  MoveL 2827 to (-200, -40.67, 52.07) mm, rotated rx 123.54 ry 0 rz 180 deg; joints [-9.323, -80.006, 124.061, 166.716, 44.832, -136.951]
  MoveL 2828 to (0, -40.67, 52.07) mm, rotated rx 123.54 ry 0 rz 180 deg; joints [-7.983, -68.226, 108.402, 167.736, 40.83, -137.116]
  MoveL 2829 to (0, -40.33, 52.56) mm, rotated rx 126.23 ry 0 rz 180 deg; joints [-8.518, -67.714, 108.589, 167.109, 41.6, -134.058]
  MoveL 2830 to (-200, -40.33, 52.56) mm, rotated rx 126.23 ry 0 rz 180 deg; joints [-9.945, -79.388, 124.274, 166.047, 45.743, -133.933]
  MoveL 2831 to (-200, -39.96, 53.04) mm, rotated rx 128.92 ry 0 rz 180 deg; joints [-10.538, -78.733, 124.49, 165.444, 46.691, -130.985]
  MoveL 2832 to (0, -39.96, 53.04) mm, rotated rx 128.92 ry 0 rz 180 deg; joints [-9.029, -67.172, 108.78, 166.542, 42.401, -131.062]
  MoveL 2833 to (0, -39.57, 53.5) mm, rotated rx 131.6 ry 0 rz 180 deg; joints [-9.515, -66.6, 108.972, 166.034, 43.23, -128.128]
  MoveL 2834 to (-200, -39.57, 53.5) mm, rotated rx 131.6 ry 0 rz 180 deg; joints [-11.101, -78.04, 124.71, 164.904, 47.673, -128.104]
  MoveL 2835 to (-200, -39.16, 53.94) mm, rotated rx 134.29 ry 0 rz 180 deg; joints [-11.634, -77.311, 124.93, 164.426, 48.684, -125.287]
  MoveL 2836 to (0, -39.16, 53.94) mm, rotated rx 134.29 ry 0 rz 180 deg; joints [-9.975, -65.998, 109.167, 165.583, 44.084, -125.251]
  MoveL 2837 to (0, -38.73, 54.36) mm, rotated rx 136.97 ry 0 rz 180 deg; joints [-10.407, -65.369, 109.361, 165.188, 44.96, -122.429]
  MoveL 2838 to (-200, -38.73, 54.36) mm, rotated rx 136.97 ry 0 rz 180 deg; joints [-12.134, -76.548, 125.152, 164.007, 49.723, -122.53]
  MoveL 2839 to (-200, -38.29, 54.76) mm, rotated rx 139.66 ry 0 rz 180 deg; joints [-12.602, -75.751, 125.373, 163.644, 50.786, -119.831]
  MoveL 2840 to (0, -38.29, 54.76) mm, rotated rx 139.66 ry 0 rz 180 deg; joints [-10.812, -64.712, 109.555, 164.846, 45.857, -119.661]
  MoveL 2841 to (0, -37.82, 55.13) mm, rotated rx 142.34 ry 0 rz 180 deg; joints [-11.188, -64.03, 109.748, 164.556, 46.771, -116.941]
  MoveL 2842 to (-200, -37.82, 55.13) mm, rotated rx 142.34 ry 0 rz 180 deg; joints [-13.037, -74.922, 125.593, 163.335, 51.871, -117.184]
  MoveL 2843 to (-200, -37.34, 55.49) mm, rotated rx 145.03 ry 0 rz 180 deg; joints [-13.438, -74.063, 125.81, 163.077, 52.974, -114.588]
  MoveL 2844 to (0, -37.34, 55.49) mm, rotated rx 145.03 ry 0 rz 180 deg; joints [-11.536, -63.323, 109.939, 164.314, 47.701, -114.267]
  MoveL 2845 to (0, -36.84, 55.82) mm, rotated rx 147.72 ry 0 rz 180 deg; joints [-11.853, -62.592, 110.127, 164.118, 48.643, -111.637]
  MoveL 2846 to (-200, -36.84, 55.82) mm, rotated rx 147.72 ry 0 rz 180 deg; joints [-13.804, -73.174, 126.025, 162.868, 54.095, -112.037]
  MoveL 2847 to (-200, -36.32, 56.13) mm, rotated rx 150.4 ry 0 rz 180 deg; joints [-14.135, -72.258, 126.235, 162.705, 55.228, -109.53]
  MoveL 2848 to (0, -36.32, 56.13) mm, rotated rx 150.4 ry 0 rz 180 deg; joints [-12.14, -61.84, 110.312, 163.968, 49.597, -109.048]
  MoveL 2849 to (0, -35.79, 56.41) mm, rotated rx 153.09 ry 0 rz 180 deg; joints [-12.397, -61.067, 110.492, 163.86, 50.559, -106.496]
  MoveL 2850 to (-200, -35.79, 56.41) mm, rotated rx 153.09 ry 0 rz 180 deg; joints [-14.43, -71.315, 126.439, 162.585, 56.374, -107.059]
  MoveL 2851 to (-200, -35.25, 56.67) mm, rotated rx 155.77 ry 0 rz 180 deg; joints [-14.69, -70.349, 126.638, 162.508, 57.53, -104.624]
  MoveL 2852 to (0, -35.25, 56.67) mm, rotated rx 155.77 ry 0 rz 180 deg; joints [-12.623, -60.276, 110.668, 163.792, 51.529, -103.977]
  MoveL 2853 to (0, -34.7, 56.91) mm, rotated rx 158.46 ry 0 rz 180 deg; joints [-12.817, -59.467, 110.837, 163.763, 52.503, -101.488]
  MoveL 2854 to (-200, -34.7, 56.91) mm, rotated rx 158.46 ry 0 rz 180 deg; joints [-14.913, -69.361, 126.83, 162.469, 58.693, -102.219]
  MoveL 2855 to (-200, -34.14, 57.11) mm, rotated rx 161.14 ry 0 rz 180 deg; joints [-15.1, -68.352, 127.015, 162.468, 59.86, -99.843]
  MoveL 2856 to (0, -34.14, 57.11) mm, rotated rx 161.14 ry 0 rz 180 deg; joints [-12.979, -58.642, 111.001, 163.771, 53.479, -99.029]
  MoveL 2857 to (0, -33.56, 57.29) mm, rotated rx 163.83 ry 0 rz 180 deg; joints [-13.11, -57.803, 111.157, 163.814, 54.458, -96.593]
  MoveL 2858 to (-200, -33.56, 57.29) mm, rotated rx 163.83 ry 0 rz 180 deg; joints [-15.25, -67.325, 127.192, 162.503, 61.031, -97.489]
  MoveL 2859 to (-200, -32.98, 57.45) mm, rotated rx 166.52 ry 0 rz 180 deg; joints [-15.363, -66.282, 127.359, 162.573, 62.203, -95.156]
  MoveL 2860 to (0, -32.98, 57.45) mm, rotated rx 166.52 ry 0 rz 180 deg; joints [-13.208, -56.951, 111.307, 163.891, 55.435, -94.179]
  MoveL 2861 to (0, -32.4, 57.57) mm, rotated rx 169.2 ry 0 rz 180 deg; joints [-13.274, -56.089, 111.449, 164, 56.411, -91.784]
  MoveL 2862 to (-200, -32.4, 57.57) mm, rotated rx 169.2 ry 0 rz 180 deg; joints [-15.439, -65.224, 127.518, 162.675, 63.374, -92.839]
  MoveL 2863 to (-200, -31.81, 57.67) mm, rotated rx 171.89 ry 0 rz 180 deg; joints [-15.478, -64.155, 127.666, 162.808, 64.542, -90.538]
  MoveL 2864 to (0, -31.81, 57.67) mm, rotated rx 171.89 ry 0 rz 180 deg; joints [-13.308, -55.218, 111.582, 164.14, 57.381, -89.406]
  MoveL 2865 to (0, -31.21, 57.74) mm, rotated rx 174.57 ry 0 rz 180 deg; joints [-13.31, -54.34, 111.707, 164.309, 58.347, -87.041]
  MoveL 2866 to (-200, -31.21, 57.74) mm, rotated rx 174.57 ry 0 rz 180 deg; joints [-15.48, -63.077, 127.805, 162.973, 65.705, -88.245]
  MoveL 2867 to (-200, -30.61, 57.78) mm, rotated rx 177.26 ry 0 rz 180 deg; joints [-15.444, -61.991, 127.932, 163.167, 66.861, -85.961]
  MoveL 2868 to (0, -30.61, 57.78) mm, rotated rx 177.26 ry 0 rz 180 deg; joints [-13.279, -53.457, 111.823, 164.508, 59.305, -84.687]
  MoveL 2869 to (0, -30.01, 57.8) mm, rotated rx 179.94 ry 0 rz 180 deg; joints [-13.215, -52.571, 111.93, 164.734, 60.254, -82.343]
  MoveL 2870 to (-200, -30.01, 57.8) mm, rotated rx 179.94 ry 0 rz 180 deg; joints [-15.371, -60.901, 128.049, 163.389, 68.009, -83.681]
  MoveL 2871 to (-200, -29.41, 57.8) mm, rotated rx 180 ry 0 rz 180 deg; joints [-15.369, -60.841, 128.054, 163.399, 68.071, -83.647]
  MoveL 2872 to (0, -29.41, 57.8) mm, rotated rx 180 ry 0 rz 180 deg; joints [-13.214, -52.522, 111.934, 164.743, 60.305, -82.305]
  MoveL 2873 to (0, -28.81, 57.8) mm, rotated rx 180 ry 0 rz 180 deg; joints [-13.214, -52.491, 111.937, 164.748, 60.337, -82.315]
  MoveL 2874 to (-200, -28.81, 57.8) mm, rotated rx 180 ry 0 rz 180 deg; joints [-15.369, -60.802, 128.056, 163.403, 68.11, -83.659]
  MoveL 2875 to (-200, -28.21, 57.8) mm, rotated rx 180 ry 0 rz 180 deg; joints [-15.369, -60.764, 128.058, 163.408, 68.149, -83.672]
  MoveL 2876 to (0, -28.21, 57.8) mm, rotated rx 180 ry 0 rz 180 deg; joints [-13.214, -52.46, 111.939, 164.753, 60.369, -82.325]
  MoveL 2877 to (0, -27.61, 57.8) mm, rotated rx 180 ry 0 rz 180 deg; joints [-13.214, -52.428, 111.941, 164.758, 60.402, -82.335]
  MoveL 2878 to (-200, -27.61, 57.8) mm, rotated rx 180 ry 0 rz 180 deg; joints [-15.369, -60.725, 128.061, 163.413, 68.188, -83.684]
  MoveL 2879 to (-200, -27.01, 57.8) mm, rotated rx 180 ry 0 rz 180 deg; joints [-15.369, -60.687, 128.063, 163.417, 68.227, -83.697]
  MoveL 2880 to (0, -27.01, 57.8) mm, rotated rx 180 ry 0 rz 180 deg; joints [-13.214, -52.397, 111.943, 164.763, 60.434, -82.345]
  MoveL 2881 to (0, -26.41, 57.8) mm, rotated rx 180 ry 0 rz 180 deg; joints [-13.214, -52.365, 111.945, 164.768, 60.466, -82.355]
  MoveL 2882 to (-200, -26.41, 57.8) mm, rotated rx 180 ry 0 rz 180 deg; joints [-15.369, -60.648, 128.065, 163.422, 68.266, -83.709]
  MoveL 2883 to (-200, -25.81, 57.8) mm, rotated rx 180 ry 0 rz 180 deg; joints [-15.369, -60.61, 128.067, 163.427, 68.306, -83.722]
  MoveL 2884 to (0, -25.81, 57.8) mm, rotated rx 180 ry 0 rz 180 deg; joints [-13.214, -52.334, 111.947, 164.773, 60.498, -82.366]
  MoveL 2885 to (0, -25.21, 57.8) mm, rotated rx 180 ry 0 rz 180 deg; joints [-13.214, -52.302, 111.949, 164.778, 60.531, -82.376]
  MoveL 2886 to (-200, -25.21, 57.8) mm, rotated rx 180 ry 0 rz 180 deg; joints [-15.369, -60.571, 128.069, 163.431, 68.345, -83.734]
  MoveL 2887 to (-200, -24.61, 57.8) mm, rotated rx 180 ry 0 rz 180 deg; joints [-15.369, -60.532, 128.071, 163.436, 68.384, -83.747]
  MoveL 2888 to (0, -24.61, 57.8) mm, rotated rx 180 ry 0 rz 180 deg; joints [-13.214, -52.271, 111.95, 164.783, 60.563, -82.386]
  MoveL 2889 to (0, -24.01, 57.8) mm, rotated rx 180 ry 0 rz 180 deg; joints [-13.214, -52.239, 111.952, 164.788, 60.595, -82.396]
  MoveL 2890 to (-200, -24.01, 57.8) mm, rotated rx 180 ry 0 rz 180 deg; joints [-15.369, -60.494, 128.073, 163.44, 68.423, -83.759]
  MoveL 2891 to (-200, -23.41, 57.8) mm, rotated rx 180 ry 0 rz 180 deg; joints [-15.369, -60.455, 128.075, 163.445, 68.462, -83.772]
  MoveL 2892 to (0, -23.41, 57.8) mm, rotated rx 180 ry 0 rz 180 deg; joints [-13.214, -52.208, 111.954, 164.793, 60.627, -82.406]
  MoveL 2893 to (0, -22.81, 57.8) mm, rotated rx 180 ry 0 rz 180 deg; joints [-13.214, -52.176, 111.956, 164.798, 60.659, -82.416]
  MoveL 2894 to (-200, -22.81, 57.8) mm, rotated rx 180 ry 0 rz 180 deg; joints [-15.369, -60.416, 128.077, 163.45, 68.501, -83.784]
  MoveL 2895 to (-200, -22.21, 57.8) mm, rotated rx 180 ry 0 rz 180 deg; joints [-15.369, -60.378, 128.079, 163.454, 68.54, -83.797]
  MoveL 2896 to (0, -22.21, 57.8) mm, rotated rx 180 ry 0 rz 180 deg; joints [-13.214, -52.145, 111.958, 164.803, 60.691, -82.426]
  MoveL 2897 to (0, -21.61, 57.8) mm, rotated rx 180 ry 0 rz 180 deg; joints [-13.214, -52.113, 111.959, 164.808, 60.724, -82.436]
  MoveL 2898 to (-200, -21.61, 57.8) mm, rotated rx 180 ry 0 rz 180 deg; joints [-15.369, -60.339, 128.081, 163.459, 68.579, -83.809]
  MoveL 2899 to (-200, -21.01, 57.8) mm, rotated rx 180 ry 0 rz 180 deg; joints [-15.369, -60.3, 128.083, 163.463, 68.618, -83.822]
  MoveL 2900 to (0, -21.01, 57.8) mm, rotated rx 180 ry 0 rz 180 deg; joints [-13.214, -52.082, 111.961, 164.813, 60.756, -82.446]
  MoveL 2901 to (0, -20.41, 57.8) mm, rotated rx 180 ry 0 rz 180 deg; joints [-13.214, -52.05, 111.963, 164.818, 60.788, -82.456]
  MoveL 2902 to (-200, -20.41, 57.8) mm, rotated rx 180 ry 0 rz 180 deg; joints [-15.369, -60.261, 128.085, 163.468, 68.657, -83.834]
  MoveL 2903 to (-200, -19.81, 57.8) mm, rotated rx 180 ry 0 rz 180 deg; joints [-15.369, -60.223, 128.087, 163.472, 68.695, -83.847]
  MoveL 2904 to (0, -19.81, 57.8) mm, rotated rx 180 ry 0 rz 180 deg; joints [-13.214, -52.018, 111.964, 164.823, 60.82, -82.466]
  MoveL 2905 to (0, -19.21, 57.8) mm, rotated rx 180 ry 0 rz 180 deg; joints [-13.214, -51.987, 111.966, 164.827, 60.852, -82.476]
  MoveL 2906 to (-200, -19.21, 57.8) mm, rotated rx 180 ry 0 rz 180 deg; joints [-15.369, -60.184, 128.089, 163.477, 68.734, -83.859]
  MoveL 2907 to (-200, -18.61, 57.8) mm, rotated rx 180 ry 0 rz 180 deg; joints [-15.369, -60.145, 128.09, 163.481, 68.773, -83.871]
  MoveL 2908 to (0, -18.61, 57.8) mm, rotated rx 180 ry 0 rz 180 deg; joints [-13.214, -51.955, 111.968, 164.832, 60.884, -82.486]
  MoveL 2909 to (0, -18.01, 57.8) mm, rotated rx 180 ry 0 rz 180 deg; joints [-13.214, -51.923, 111.969, 164.837, 60.916, -82.496]
  MoveL 2910 to (-200, -18.01, 57.8) mm, rotated rx 180 ry 0 rz 180 deg; joints [-15.369, -60.106, 128.092, 163.486, 68.812, -83.884]
  MoveL 2911 to (-200, -17.41, 57.8) mm, rotated rx 180 ry 0 rz 180 deg; joints [-15.369, -60.067, 128.094, 163.49, 68.851, -83.896]
  MoveL 2912 to (0, -17.41, 57.8) mm, rotated rx 180 ry 0 rz 180 deg; joints [-13.214, -51.892, 111.971, 164.842, 60.948, -82.506]
  MoveL 2913 to (0, -16.81, 57.8) mm, rotated rx 180 ry 0 rz 180 deg; joints [-13.214, -51.86, 111.972, 164.847, 60.98, -82.516]
  MoveL 2914 to (-200, -16.81, 57.8) mm, rotated rx 180 ry 0 rz 180 deg; joints [-15.369, -60.028, 128.096, 163.495, 68.89, -83.908]
  MoveL 2915 to (-200, -16.21, 57.8) mm, rotated rx 180 ry 0 rz 180 deg; joints [-15.369, -59.989, 128.097, 163.499, 68.929, -83.921]
  MoveL 2916 to (0, -16.21, 57.8) mm, rotated rx 180 ry 0 rz 180 deg; joints [-13.214, -51.828, 111.974, 164.852, 61.012, -82.525]
  MoveL 2917 to (0, -15.61, 57.8) mm, rotated rx 180 ry 0 rz 180 deg; joints [-13.214, -51.797, 111.975, 164.856, 61.044, -82.535]
  MoveL 2918 to (-200, -15.61, 57.8) mm, rotated rx 180 ry 0 rz 180 deg; joints [-15.369, -59.95, 128.099, 163.503, 68.968, -83.933]
  MoveL 2919 to (-200, -15.01, 57.8) mm, rotated rx 180 ry 0 rz 180 deg; joints [-15.369, -59.912, 128.1, 163.508, 69.006, -83.945]
  MoveL 2920 to (0, -15.01, 57.8) mm, rotated rx 180 ry 0 rz 180 deg; joints [-13.214, -51.765, 111.976, 164.861, 61.076, -82.545]
  MoveL 2921 to (0, -14.41, 57.8) mm, rotated rx 180 ry 0 rz 180 deg; joints [-13.214, -51.733, 111.978, 164.866, 61.108, -82.555]
  MoveL 2922 to (-200, -14.41, 57.8) mm, rotated rx 180 ry 0 rz 180 deg; joints [-15.369, -59.873, 128.102, 163.512, 69.045, -83.958]
  MoveL 2923 to (-200, -13.81, 57.8) mm, rotated rx 180 ry 0 rz 180 deg; joints [-15.369, -59.834, 128.103, 163.517, 69.084, -83.97]
  MoveL 2924 to (0, -13.81, 57.8) mm, rotated rx 180 ry 0 rz 180 deg; joints [-13.214, -51.701, 111.979, 164.871, 61.14, -82.565]
  MoveL 2925 to (0, -13.21, 57.8) mm, rotated rx 180 ry 0 rz 180 deg; joints [-13.214, -51.67, 111.981, 164.875, 61.172, -82.575]
  MoveL 2926 to (-200, -13.21, 57.8) mm, rotated rx 180 ry 0 rz 180 deg; joints [-15.369, -59.795, 128.105, 163.521, 69.123, -83.982]
  MoveL 2927 to (-200, -12.61, 57.8) mm, rotated rx 180 ry 0 rz 180 deg; joints [-15.369, -59.756, 128.106, 163.525, 69.162, -83.994]
  MoveL 2928 to (0, -12.61, 57.8) mm, rotated rx 180 ry 0 rz 180 deg; joints [-13.214, -51.638, 111.982, 164.88, 61.204, -82.585]
  MoveL 2929 to (0, -12.01, 57.8) mm, rotated rx 180 ry 0 rz 180 deg; joints [-13.214, -51.606, 111.983, 164.885, 61.236, -82.595]
  MoveL 2930 to (-200, -12.01, 57.8) mm, rotated rx 180 ry 0 rz 180 deg; joints [-15.369, -59.717, 128.108, 163.53, 69.2, -84.007]
  MoveL 2931 to (-200, -11.41, 57.8) mm, rotated rx 180 ry 0 rz 180 deg; joints [-15.369, -59.678, 128.109, 163.534, 69.239, -84.019]
  MoveL 2932 to (0, -11.41, 57.8) mm, rotated rx 180 ry 0 rz 180 deg; joints [-13.214, -51.574, 111.984, 164.89, 61.268, -82.604]
  MoveL 2933 to (0, -10.81, 57.8) mm, rotated rx 180 ry 0 rz 180 deg; joints [-13.214, -51.542, 111.985, 164.894, 61.3, -82.614]
  MoveL 2934 to (-200, -10.81, 57.8) mm, rotated rx 180 ry 0 rz 180 deg; joints [-15.369, -59.639, 128.11, 163.538, 69.278, -84.031]
  MoveL 2935 to (-200, -10.21, 57.8) mm, rotated rx 180 ry 0 rz 180 deg; joints [-15.369, -59.599, 128.112, 163.543, 69.317, -84.043]
  MoveL 2936 to (0, -10.21, 57.8) mm, rotated rx 180 ry 0 rz 180 deg; joints [-13.214, -51.51, 111.987, 164.899, 61.332, -82.624]
  MoveL 2937 to (0, -9.61, 57.8) mm, rotated rx 180 ry 0 rz 180 deg; joints [-13.214, -51.478, 111.988, 164.904, 61.364, -82.634]
  MoveL 2938 to (-200, -9.61, 57.8) mm, rotated rx 180 ry 0 rz 180 deg; joints [-15.369, -59.56, 128.113, 163.547, 69.355, -84.056]
  MoveL 2939 to (-200, -9.01, 57.8) mm, rotated rx 180 ry 0 rz 180 deg; joints [-15.369, -59.521, 128.114, 163.551, 69.394, -84.068]
  MoveL 2940 to (0, -9.01, 57.8) mm, rotated rx 180 ry 0 rz 180 deg; joints [-13.214, -51.447, 111.989, 164.908, 61.396, -82.644]
  MoveL 2941 to (0, -8.41, 57.8) mm, rotated rx 180 ry 0 rz 180 deg; joints [-13.214, -51.415, 111.99, 164.913, 61.427, -82.653]
  MoveL 2942 to (-200, -8.41, 57.8) mm, rotated rx 180 ry 0 rz 180 deg; joints [-15.369, -59.482, 128.115, 163.556, 69.433, -84.08]
  MoveL 2943 to (-200, -7.81, 57.8) mm, rotated rx 180 ry 0 rz 180 deg; joints [-15.369, -59.443, 128.116, 163.56, 69.471, -84.092]
  MoveL 2944 to (0, -7.81, 57.8) mm, rotated rx 180 ry 0 rz 180 deg; joints [-13.214, -51.383, 111.991, 164.918, 61.459, -82.663]
  MoveL 2945 to (0, -7.21, 57.8) mm, rotated rx 180 ry 0 rz 180 deg; joints [-13.214, -51.351, 111.992, 164.922, 61.491, -82.673]
  MoveL 2946 to (-200, -7.21, 57.8) mm, rotated rx 180 ry 0 rz 180 deg; joints [-15.369, -59.404, 128.118, 163.564, 69.51, -84.104]
  MoveL 2947 to (-200, -6.61, 57.8) mm, rotated rx 180 ry 0 rz 180 deg; joints [-15.369, -59.365, 128.119, 163.568, 69.549, -84.117]
  MoveL 2948 to (0, -6.61, 57.8) mm, rotated rx 180 ry 0 rz 180 deg; joints [-13.214, -51.319, 111.993, 164.927, 61.523, -82.683]
  MoveL 2949 to (0, -6.01, 57.8) mm, rotated rx 180 ry 0 rz 180 deg; joints [-13.214, -51.287, 111.994, 164.932, 61.555, -82.692]
  MoveL 2950 to (-200, -6.01, 57.8) mm, rotated rx 180 ry 0 rz 180 deg; joints [-15.369, -59.326, 128.12, 163.573, 69.587, -84.129]
  MoveL 2951 to (-200, -5.41, 57.8) mm, rotated rx 180 ry 0 rz 180 deg; joints [-15.369, -59.286, 128.121, 163.577, 69.626, -84.141]
  MoveL 2952 to (0, -5.41, 57.8) mm, rotated rx 180 ry 0 rz 180 deg; joints [-13.214, -51.255, 111.995, 164.936, 61.587, -82.702]
  MoveL 2953 to (0, -4.81, 57.8) mm, rotated rx 180 ry 0 rz 180 deg; joints [-13.214, -51.223, 111.996, 164.941, 61.618, -82.712]
  MoveL 2954 to (-200, -4.81, 57.8) mm, rotated rx 180 ry 0 rz 180 deg; joints [-15.369, -59.247, 128.122, 163.581, 69.664, -84.153]
  MoveL 2955 to (-200, -4.21, 57.8) mm, rotated rx 180 ry 0 rz 180 deg; joints [-15.369, -59.208, 128.123, 163.585, 69.703, -84.165]
  MoveL 2956 to (0, -4.21, 57.8) mm, rotated rx 180 ry 0 rz 180 deg; joints [-13.214, -51.191, 111.997, 164.946, 61.65, -82.722]
  MoveL 2957 to (0, -3.61, 57.8) mm, rotated rx 180 ry 0 rz 180 deg; joints [-13.214, -51.159, 111.998, 164.95, 61.682, -82.731]
  MoveL 2958 to (-200, -3.61, 57.8) mm, rotated rx 180 ry 0 rz 180 deg; joints [-15.369, -59.169, 128.124, 163.59, 69.741, -84.177]
  MoveL 2959 to (-200, -3.01, 57.8) mm, rotated rx 180 ry 0 rz 180 deg; joints [-15.369, -59.129, 128.125, 163.594, 69.78, -84.189]
  MoveL 2960 to (0, -3.01, 57.8) mm, rotated rx 180 ry 0 rz 180 deg; joints [-13.214, -51.127, 111.998, 164.955, 61.714, -82.741]
  MoveL 2961 to (0, -2.41, 57.8) mm, rotated rx 180 ry 0 rz 180 deg; joints [-13.214, -51.095, 111.999, 164.959, 61.745, -82.751]
  MoveL 2962 to (-200, -2.41, 57.8) mm, rotated rx 180 ry 0 rz 180 deg; joints [-15.369, -59.09, 128.125, 163.598, 69.819, -84.201]
  MoveL 2963 to (-200, -1.81, 57.8) mm, rotated rx 180 ry 0 rz 180 deg; joints [-15.369, -59.051, 128.126, 163.602, 69.857, -84.213]
  MoveL 2964 to (0, -1.81, 57.8) mm, rotated rx 180 ry 0 rz 180 deg; joints [-13.214, -51.063, 112, 164.964, 61.777, -82.76]
  MoveL 2965 to (0, -1.21, 57.8) mm, rotated rx 180 ry 0 rz 180 deg; joints [-13.214, -51.03, 112.001, 164.969, 61.809, -82.77]
  MoveL 2966 to (-200, -1.21, 57.8) mm, rotated rx 180 ry 0 rz 180 deg; joints [-15.369, -59.011, 128.127, 163.606, 69.896, -84.226]
  MoveL 2967 to (-200, -0.61, 57.8) mm, rotated rx 180 ry 0 rz 180 deg; joints [-15.369, -58.972, 128.128, 163.61, 69.934, -84.238]
  MoveL 2968 to (0, -0.61, 57.8) mm, rotated rx 180 ry 0 rz 180 deg; joints [-13.214, -50.998, 112.001, 164.973, 61.84, -82.78]
  MoveL 2969 to (0, -0.01, 57.8) mm, rotated rx 180 ry 0 rz 180 deg; joints [-13.214, -50.966, 112.002, 164.978, 61.872, -82.789]
  MoveL 2970 to (-200, -0.01, 57.8) mm, rotated rx 180 ry 0 rz 180 deg; joints [-15.369, -58.933, 128.129, 163.614, 69.972, -84.25]
  MoveL 2971 to (-200, 0, 57.8) mm, rotated rx 180 ry 0 rz 180 deg; joints [-15.369, -58.932, 128.129, 163.615, 69.973, -84.25]
  MoveL 2972 to (0, 0, 57.8) mm, rotated rx 180 ry 0 rz 180 deg; joints [-13.214, -50.966, 112.002, 164.978, 61.873, -82.789]
  MoveL 2973 to (0, 0, 58.2) mm, rotated rx 180 ry 0 rz 180 deg; joints [-13.23, -50.962, 111.994, 164.959, 61.871, -82.78]
  MoveL 2974 to (-200, 0, 58.2) mm, rotated rx 180 ry 0 rz 180 deg; joints [-15.388, -58.928, 128.12, 163.595, 69.971, -84.242]
  MoveL 2975 to (-200, -0.6, 58.2) mm, rotated rx 180 ry 0 rz 180 deg; joints [-15.388, -58.967, 128.119, 163.591, 69.933, -84.23]
  MoveL 2976 to (0, -0.6, 58.2) mm, rotated rx 180 ry 0 rz 180 deg; joints [-13.23, -50.994, 111.993, 164.955, 61.839, -82.77]
  MoveL 2977 to (0, -1.2, 58.2) mm, rotated rx 180 ry 0 rz 180 deg; joints [-13.23, -51.026, 111.993, 164.95, 61.807, -82.761]
  MoveL 2978 to (-200, -1.2, 58.2) mm, rotated rx 180 ry 0 rz 180 deg; joints [-15.388, -59.006, 128.119, 163.587, 69.894, -84.218]
  MoveL 2979 to (-200, -1.8, 58.2) mm, rotated rx 180 ry 0 rz 180 deg; joints [-15.388, -59.046, 128.118, 163.582, 69.856, -84.206]
  MoveL 2980 to (0, -1.8, 58.2) mm, rotated rx 180 ry 0 rz 180 deg; joints [-13.23, -51.058, 111.992, 164.946, 61.776, -82.751]
  MoveL 2981 to (0, -2.4, 58.2) mm, rotated rx 180 ry 0 rz 180 deg; joints [-13.23, -51.09, 111.991, 164.941, 61.744, -82.741]
  MoveL 2982 to (-200, -2.4, 58.2) mm, rotated rx 180 ry 0 rz 180 deg; joints [-15.388, -59.085, 128.117, 163.578, 69.817, -84.194]
  MoveL 2983 to (-200, -3, 58.2) mm, rotated rx 180 ry 0 rz 180 deg; joints [-15.388, -59.124, 128.116, 163.574, 69.779, -84.182]
  MoveL 2984 to (0, -3, 58.2) mm, rotated rx 180 ry 0 rz 180 deg; joints [-13.23, -51.122, 111.99, 164.937, 61.712, -82.732]
  MoveL 2985 to (0, -3.6, 58.2) mm, rotated rx 180 ry 0 rz 180 deg; joints [-13.23, -51.154, 111.99, 164.932, 61.681, -82.722]
  MoveL 2986 to (-200, -3.6, 58.2) mm, rotated rx 180 ry 0 rz 180 deg; joints [-15.388, -59.164, 128.115, 163.57, 69.74, -84.17]
  MoveL 2987 to (-200, -4.2, 58.2) mm, rotated rx 180 ry 0 rz 180 deg; joints [-15.388, -59.203, 128.114, 163.566, 69.701, -84.157]
  MoveL 2988 to (0, -4.2, 58.2) mm, rotated rx 180 ry 0 rz 180 deg; joints [-13.23, -51.186, 111.989, 164.927, 61.649, -82.712]
  MoveL 2989 to (0, -4.8, 58.2) mm, rotated rx 180 ry 0 rz 180 deg; joints [-13.23, -51.218, 111.988, 164.923, 61.617, -82.702]
  MoveL 2990 to (-200, -4.8, 58.2) mm, rotated rx 180 ry 0 rz 180 deg; joints [-15.388, -59.242, 128.113, 163.561, 69.663, -84.145]
  MoveL 2991 to (-200, -5.4, 58.2) mm, rotated rx 180 ry 0 rz 180 deg; joints [-15.388, -59.281, 128.112, 163.557, 69.624, -84.133]
  MoveL 2992 to (0, -5.4, 58.2) mm, rotated rx 180 ry 0 rz 180 deg; joints [-13.23, -51.25, 111.987, 164.918, 61.585, -82.693]
  MoveL 2993 to (0, -6, 58.2) mm, rotated rx 180 ry 0 rz 180 deg; joints [-13.23, -51.282, 111.986, 164.913, 61.553, -82.683]
  MoveL 2994 to (-200, -6, 58.2) mm, rotated rx 180 ry 0 rz 180 deg; joints [-15.388, -59.321, 128.111, 163.553, 69.586, -84.121]
  MoveL 2995 to (-200, -6.6, 58.2) mm, rotated rx 180 ry 0 rz 180 deg; joints [-15.388, -59.36, 128.11, 163.549, 69.547, -84.109]
  MoveL 2996 to (0, -6.6, 58.2) mm, rotated rx 180 ry 0 rz 180 deg; joints [-13.23, -51.314, 111.985, 164.909, 61.522, -82.673]
  MoveL 2997 to (0, -7.2, 58.2) mm, rotated rx 180 ry 0 rz 180 deg; joints [-13.23, -51.346, 111.984, 164.904, 61.49, -82.663]
  MoveL 2998 to (-200, -7.2, 58.2) mm, rotated rx 180 ry 0 rz 180 deg; joints [-15.388, -59.399, 128.109, 163.545, 69.509, -84.097]
  MoveL 2999 to (-200, -7.8, 58.2) mm, rotated rx 180 ry 0 rz 180 deg; joints [-15.388, -59.438, 128.108, 163.54, 69.47, -84.084]
  MoveL 3000 to (0, -7.8, 58.2) mm, rotated rx 180 ry 0 rz 180 deg; joints [-13.23, -51.378, 111.983, 164.899, 61.458, -82.654]
  MoveL 3001 to (0, -8.4, 58.2) mm, rotated rx 180 ry 0 rz 180 deg; joints [-13.23, -51.41, 111.982, 164.895, 61.426, -82.644]
  MoveL 3002 to (-200, -8.4, 58.2) mm, rotated rx 180 ry 0 rz 180 deg; joints [-15.388, -59.477, 128.107, 163.536, 69.431, -84.072]
  MoveL 3003 to (-200, -9, 58.2) mm, rotated rx 180 ry 0 rz 180 deg; joints [-15.388, -59.516, 128.106, 163.532, 69.393, -84.06]
  MoveL 3004 to (0, -9, 58.2) mm, rotated rx 180 ry 0 rz 180 deg; joints [-13.23, -51.442, 111.981, 164.89, 61.394, -82.634]
  MoveL 3005 to (0, -9.6, 58.2) mm, rotated rx 180 ry 0 rz 180 deg; joints [-13.23, -51.474, 111.98, 164.885, 61.363, -82.624]
  MoveL 3006 to (-200, -9.6, 58.2) mm, rotated rx 180 ry 0 rz 180 deg; joints [-15.388, -59.555, 128.104, 163.527, 69.354, -84.048]
  MoveL 3007 to (-200, -10.2, 58.2) mm, rotated rx 180 ry 0 rz 180 deg; joints [-15.388, -59.594, 128.103, 163.523, 69.315, -84.036]
  MoveL 3008 to (0, -10.2, 58.2) mm, rotated rx 180 ry 0 rz 180 deg; joints [-13.23, -51.506, 111.979, 164.881, 61.331, -82.614]
  MoveL 3009 to (0, -10.8, 58.2) mm, rotated rx 180 ry 0 rz 180 deg; joints [-13.23, -51.538, 111.978, 164.876, 61.299, -82.605]
  MoveL 3010 to (-200, -10.8, 58.2) mm, rotated rx 180 ry 0 rz 180 deg; joints [-15.388, -59.634, 128.102, 163.519, 69.276, -84.023]
  MoveL 3011 to (-200, -11.4, 58.2) mm, rotated rx 180 ry 0 rz 180 deg; joints [-15.388, -59.673, 128.101, 163.514, 69.238, -84.011]
  MoveL 3012 to (0, -11.4, 58.2) mm, rotated rx 180 ry 0 rz 180 deg; joints [-13.23, -51.569, 111.976, 164.871, 61.267, -82.595]
  MoveL 3013 to (0, -12, 58.2) mm, rotated rx 180 ry 0 rz 180 deg; joints [-13.23, -51.601, 111.975, 164.867, 61.235, -82.585]
  MoveL 3014 to (-200, -12, 58.2) mm, rotated rx 180 ry 0 rz 180 deg; joints [-15.388, -59.712, 128.099, 163.51, 69.199, -83.999]
  MoveL 3015 to (-200, -12.6, 58.2) mm, rotated rx 180 ry 0 rz 180 deg; joints [-15.388, -59.751, 128.098, 163.506, 69.16, -83.987]
  MoveL 3016 to (0, -12.6, 58.2) mm, rotated rx 180 ry 0 rz 180 deg; joints [-13.23, -51.633, 111.974, 164.862, 61.203, -82.575]
  MoveL 3017 to (0, -13.2, 58.2) mm, rotated rx 180 ry 0 rz 180 deg; joints [-13.23, -51.665, 111.973, 164.857, 61.171, -82.565]
  MoveL 3018 to (-200, -13.2, 58.2) mm, rotated rx 180 ry 0 rz 180 deg; joints [-15.388, -59.79, 128.096, 163.501, 69.122, -83.974]
  MoveL 3019 to (-200, -13.8, 58.2) mm, rotated rx 180 ry 0 rz 180 deg; joints [-15.388, -59.829, 128.095, 163.497, 69.083, -83.962]
  MoveL 3020 to (0, -13.8, 58.2) mm, rotated rx 180 ry 0 rz 180 deg; joints [-13.23, -51.697, 111.971, 164.852, 61.139, -82.555]
  MoveL 3021 to (0, -14.4, 58.2) mm, rotated rx 180 ry 0 rz 180 deg; joints [-13.23, -51.728, 111.97, 164.847, 61.107, -82.545]
  MoveL 3022 to (-200, -14.4, 58.2) mm, rotated rx 180 ry 0 rz 180 deg; joints [-15.388, -59.868, 128.093, 163.493, 69.044, -83.95]
  MoveL 3023 to (-200, -15, 58.2) mm, rotated rx 180 ry 0 rz 180 deg; joints [-15.388, -59.907, 128.092, 163.488, 69.005, -83.937]
  MoveL 3024 to (0, -15, 58.2) mm, rotated rx 180 ry 0 rz 180 deg; joints [-13.23, -51.76, 111.968, 164.843, 61.075, -82.536]
  MoveL 3025 to (0, -15.6, 58.2) mm, rotated rx 180 ry 0 rz 180 deg; joints [-13.23, -51.792, 111.967, 164.838, 61.043, -82.526]
  MoveL 3026 to (-200, -15.6, 58.2) mm, rotated rx 180 ry 0 rz 180 deg; joints [-15.388, -59.945, 128.09, 163.484, 68.966, -83.925]
  MoveL 3027 to (-200, -16.2, 58.2) mm, rotated rx 180 ry 0 rz 180 deg; joints [-15.388, -59.984, 128.089, 163.479, 68.928, -83.913]
  MoveL 3028 to (0, -16.2, 58.2) mm, rotated rx 180 ry 0 rz 180 deg; joints [-13.23, -51.824, 111.966, 164.833, 61.011, -82.516]
  MoveL 3029 to (0, -16.8, 58.2) mm, rotated rx 180 ry 0 rz 180 deg; joints [-13.23, -51.855, 111.964, 164.828, 60.979, -82.506]
  MoveL 3030 to (-200, -16.8, 58.2) mm, rotated rx 180 ry 0 rz 180 deg; joints [-15.388, -60.023, 128.087, 163.475, 68.889, -83.9]
  MoveL 3031 to (-200, -17.4, 58.2) mm, rotated rx 180 ry 0 rz 180 deg; joints [-15.388, -60.062, 128.085, 163.47, 68.85, -83.888]
  MoveL 3032 to (0, -17.4, 58.2) mm, rotated rx 180 ry 0 rz 180 deg; joints [-13.23, -51.887, 111.963, 164.823, 60.947, -82.496]
  MoveL 3033 to (0, -18, 58.2) mm, rotated rx 180 ry 0 rz 180 deg; joints [-13.23, -51.919, 111.961, 164.819, 60.915, -82.486]
  MoveL 3034 to (-200, -18, 58.2) mm, rotated rx 180 ry 0 rz 180 deg; joints [-15.388, -60.101, 128.084, 163.466, 68.811, -83.876]
  MoveL 3035 to (-200, -18.6, 58.2) mm, rotated rx 180 ry 0 rz 180 deg; joints [-15.388, -60.14, 128.082, 163.461, 68.772, -83.863]
  MoveL 3036 to (0, -18.6, 58.2) mm, rotated rx 180 ry 0 rz 180 deg; joints [-13.23, -51.95, 111.96, 164.814, 60.883, -82.476]
  MoveL 3037 to (0, -19.2, 58.2) mm, rotated rx 180 ry 0 rz 180 deg; joints [-13.23, -51.982, 111.958, 164.809, 60.851, -82.466]
  MoveL 3038 to (-200, -19.2, 58.2) mm, rotated rx 180 ry 0 rz 180 deg; joints [-15.388, -60.179, 128.08, 163.457, 68.733, -83.851]
  MoveL 3039 to (-200, -19.8, 58.2) mm, rotated rx 180 ry 0 rz 180 deg; joints [-15.388, -60.217, 128.079, 163.452, 68.694, -83.838]
  MoveL 3040 to (0, -19.8, 58.2) mm, rotated rx 180 ry 0 rz 180 deg; joints [-13.23, -52.014, 111.956, 164.804, 60.819, -82.456]
  MoveL 3041 to (0, -20.4, 58.2) mm, rotated rx 180 ry 0 rz 180 deg; joints [-13.23, -52.045, 111.955, 164.799, 60.787, -82.446]
  MoveL 3042 to (-200, -20.4, 58.2) mm, rotated rx 180 ry 0 rz 180 deg; joints [-15.388, -60.256, 128.077, 163.448, 68.655, -83.826]
  MoveL 3043 to (-200, -21, 58.2) mm, rotated rx 180 ry 0 rz 180 deg; joints [-15.388, -60.295, 128.075, 163.443, 68.616, -83.814]
  MoveL 3044 to (0, -21, 58.2) mm, rotated rx 180 ry 0 rz 180 deg; joints [-13.23, -52.077, 111.953, 164.794, 60.755, -82.436]
  MoveL 3045 to (0, -21.6, 58.2) mm, rotated rx 180 ry 0 rz 180 deg; joints [-13.23, -52.108, 111.951, 164.789, 60.722, -82.426]
  MoveL 3046 to (-200, -21.6, 58.2) mm, rotated rx 180 ry 0 rz 180 deg; joints [-15.388, -60.334, 128.073, 163.439, 68.577, -83.801]
  MoveL 3047 to (-200, -22.2, 58.2) mm, rotated rx 180 ry 0 rz 180 deg; joints [-15.388, -60.372, 128.071, 163.434, 68.538, -83.789]
  MoveL 3048 to (0, -22.2, 58.2) mm, rotated rx 180 ry 0 rz 180 deg; joints [-13.23, -52.14, 111.95, 164.785, 60.69, -82.416]
  MoveL 3049 to (0, -22.8, 58.2) mm, rotated rx 180 ry 0 rz 180 deg; joints [-13.23, -52.172, 111.948, 164.78, 60.658, -82.406]
  MoveL 3050 to (-200, -22.8, 58.2) mm, rotated rx 180 ry 0 rz 180 deg; joints [-15.388, -60.411, 128.069, 163.43, 68.5, -83.776]
  MoveL 3051 to (-200, -23.4, 58.2) mm, rotated rx 180 ry 0 rz 180 deg; joints [-15.388, -60.45, 128.067, 163.425, 68.461, -83.764]
  MoveL 3052 to (0, -23.4, 58.2) mm, rotated rx 180 ry 0 rz 180 deg; joints [-13.23, -52.203, 111.946, 164.775, 60.626, -82.396]
  MoveL 3053 to (0, -24, 58.2) mm, rotated rx 180 ry 0 rz 180 deg; joints [-13.23, -52.235, 111.944, 164.77, 60.594, -82.386]
  MoveL 3054 to (-200, -24, 58.2) mm, rotated rx 180 ry 0 rz 180 deg; joints [-15.388, -60.489, 128.065, 163.421, 68.422, -83.751]
  MoveL 3055 to (-200, -24.6, 58.2) mm, rotated rx 180 ry 0 rz 180 deg; joints [-15.388, -60.527, 128.063, 163.416, 68.382, -83.739]
  MoveL 3056 to (0, -24.6, 58.2) mm, rotated rx 180 ry 0 rz 180 deg; joints [-13.23, -52.266, 111.942, 164.765, 60.562, -82.376]
  MoveL 3057 to (0, -25.2, 58.2) mm, rotated rx 180 ry 0 rz 180 deg; joints [-13.23, -52.298, 111.941, 164.76, 60.529, -82.366]
  MoveL 3058 to (-200, -25.2, 58.2) mm, rotated rx 180 ry 0 rz 180 deg; joints [-15.388, -60.566, 128.061, 163.411, 68.343, -83.726]
  MoveL 3059 to (-200, -25.8, 58.2) mm, rotated rx 180 ry 0 rz 180 deg; joints [-15.388, -60.604, 128.059, 163.407, 68.304, -83.714]
  MoveL 3060 to (0, -25.8, 58.2) mm, rotated rx 180 ry 0 rz 180 deg; joints [-13.23, -52.329, 111.939, 164.755, 60.497, -82.356]
  MoveL 3061 to (0, -26.4, 58.2) mm, rotated rx 180 ry 0 rz 180 deg; joints [-13.23, -52.361, 111.937, 164.75, 60.465, -82.346]
  MoveL 3062 to (-200, -26.4, 58.2) mm, rotated rx 180 ry 0 rz 180 deg; joints [-15.388, -60.643, 128.057, 163.402, 68.265, -83.701]
  MoveL 3063 to (-200, -27, 58.2) mm, rotated rx 180 ry 0 rz 180 deg; joints [-15.388, -60.682, 128.054, 163.397, 68.226, -83.689]
  MoveL 3064 to (0, -27, 58.2) mm, rotated rx 180 ry 0 rz 180 deg; joints [-13.23, -52.392, 111.935, 164.745, 60.433, -82.335]
  MoveL 3065 to (0, -27.6, 58.2) mm, rotated rx 180 ry 0 rz 180 deg; joints [-13.23, -52.423, 111.933, 164.74, 60.401, -82.325]
  MoveL 3066 to (-200, -27.6, 58.2) mm, rotated rx 180 ry 0 rz 180 deg; joints [-15.388, -60.72, 128.052, 163.393, 68.187, -83.676]
  MoveL 3067 to (-200, -28.2, 58.2) mm, rotated rx 180 ry 0 rz 180 deg; joints [-15.388, -60.759, 128.05, 163.388, 68.148, -83.664]
  MoveL 3068 to (0, -28.2, 58.2) mm, rotated rx 180 ry 0 rz 180 deg; joints [-13.23, -52.455, 111.931, 164.735, 60.368, -82.315]
  MoveL 3069 to (0, -28.8, 58.2) mm, rotated rx 180 ry 0 rz 180 deg; joints [-13.23, -52.486, 111.929, 164.73, 60.336, -82.305]
  MoveL 3070 to (-200, -28.8, 58.2) mm, rotated rx 180 ry 0 rz 180 deg; joints [-15.388, -60.797, 128.048, 163.383, 68.109, -83.651]
  MoveL 3071 to (-200, -29.4, 58.2) mm, rotated rx 180 ry 0 rz 180 deg; joints [-15.388, -60.836, 128.045, 163.379, 68.07, -83.638]
  MoveL 3072 to (0, -29.4, 58.2) mm, rotated rx 180 ry 0 rz 180 deg; joints [-13.23, -52.518, 111.927, 164.725, 60.304, -82.295]
  MoveL 3073 to (0, -30, 58.2) mm, rotated rx 180 ry 0 rz 180 deg; joints [-13.23, -52.549, 111.924, 164.72, 60.271, -82.285]
  MoveL 3074 to (-200, -30, 58.2) mm, rotated rx 180 ry 0 rz 180 deg; joints [-15.388, -60.874, 128.043, 163.374, 68.031, -83.626]
  MoveL 3075 to (-200, -30.6, 58.19) mm, rotated rx 177.4 ry 0 rz 180 deg; joints [-15.459, -61.932, 127.93, 163.157, 66.917, -85.835]
  MoveL 3076 to (0, -30.6, 58.19) mm, rotated rx 177.4 ry 0 rz 180 deg; joints [-13.292, -53.409, 111.821, 164.499, 59.351, -84.557]
  MoveL 3077 to (0, -31.2, 58.15) mm, rotated rx 174.79 ry 0 rz 180 deg; joints [-13.324, -54.266, 111.708, 164.305, 58.422, -86.838]
  MoveL 3078 to (-200, -31.2, 58.15) mm, rotated rx 174.79 ry 0 rz 180 deg; joints [-15.496, -62.987, 127.807, 162.967, 65.795, -88.05]
  MoveL 3079 to (-200, -31.79, 58.08) mm, rotated rx 172.19 ry 0 rz 180 deg; joints [-15.498, -64.034, 127.673, 162.805, 64.667, -90.27]
  MoveL 3080 to (0, -31.79, 58.08) mm, rotated rx 172.19 ry 0 rz 180 deg; joints [-13.326, -55.119, 111.588, 164.137, 57.485, -89.129]
  MoveL 3081 to (0, -32.39, 57.98) mm, rotated rx 169.58 ry 0 rz 180 deg; joints [-13.297, -55.965, 111.459, 163.998, 56.544, -91.433]
  MoveL 3082 to (-200, -32.39, 57.98) mm, rotated rx 169.58 ry 0 rz 180 deg; joints [-15.465, -65.073, 127.53, 162.671, 63.534, -92.5]
  MoveL 3083 to (-200, -32.97, 57.86) mm, rotated rx 166.98 ry 0 rz 180 deg; joints [-15.397, -66.101, 127.378, 162.567, 62.398, -94.744]
  MoveL 3084 to (0, -32.97, 57.86) mm, rotated rx 166.98 ry 0 rz 180 deg; joints [-13.237, -56.804, 111.323, 163.887, 55.597, -93.752]
  MoveL 3085 to (0, -33.56, 57.71) mm, rotated rx 164.37 ry 0 rz 180 deg; joints [-13.148, -57.632, 111.179, 163.807, 54.649, -96.088]
  MoveL 3086 to (-200, -33.56, 57.71) mm, rotated rx 164.37 ry 0 rz 180 deg; joints [-15.293, -67.116, 127.217, 162.493, 61.261, -97.002]
  MoveL 3087 to (-200, -34.13, 57.54) mm, rotated rx 161.77 ry 0 rz 180 deg; joints [-15.156, -68.116, 127.047, 162.452, 60.124, -99.278]
  MoveL 3088 to (0, -34.13, 57.54) mm, rotated rx 161.77 ry 0 rz 180 deg; joints [-13.028, -58.449, 111.029, 163.757, 53.7, -98.444]
  MoveL 3089 to (0, -34.7, 57.34) mm, rotated rx 159.16 ry 0 rz 180 deg; joints [-12.878, -59.253, 110.872, 163.741, 52.751, -100.824]
  MoveL 3090 to (-200, -34.7, 57.34) mm, rotated rx 159.16 ry 0 rz 180 deg; joints [-14.983, -69.1, 126.87, 162.443, 58.99, -101.577]
  MoveL 3091 to (-200, -35.25, 57.11) mm, rotated rx 156.56 ry 0 rz 180 deg; joints [-14.776, -70.065, 126.685, 162.47, 57.86, -103.9]
  MoveL 3092 to (0, -35.25, 57.11) mm, rotated rx 156.56 ry 0 rz 180 deg; joints [-12.698, -60.043, 110.708, 163.759, 51.805, -103.228]
  MoveL 3093 to (0, -35.8, 56.86) mm, rotated rx 153.96 ry 0 rz 180 deg; joints [-12.488, -60.817, 110.54, 163.812, 50.862, -105.661]
  MoveL 3094 to (-200, -35.8, 56.86) mm, rotated rx 153.96 ry 0 rz 180 deg; joints [-14.535, -71.01, 126.494, 162.533, 56.736, -106.252]
  MoveL 3095 to (-200, -36.33, 56.58) mm, rotated rx 151.35 ry 0 rz 180 deg; joints [-14.26, -71.932, 126.297, 162.635, 55.621, -108.634]
  MoveL 3096 to (0, -36.33, 56.58) mm, rotated rx 151.35 ry 0 rz 180 deg; joints [-12.249, -61.573, 110.366, 163.904, 49.926, -108.124]
  MoveL 3097 to (0, -36.85, 56.28) mm, rotated rx 148.75 ry 0 rz 180 deg; joints [-11.981, -62.311, 110.188, 164.034, 48.997, -110.621]
  MoveL 3098 to (-200, -36.85, 56.28) mm, rotated rx 148.75 ry 0 rz 180 deg; joints [-13.951, -72.831, 126.095, 162.777, 54.515, -111.051]
  MoveL 3099 to (-200, -37.35, 55.96) mm, rotated rx 146.14 ry 0 rz 180 deg; joints [-13.609, -73.705, 125.888, 162.962, 53.422, -113.508]
  MoveL 3100 to (0, -37.35, 55.96) mm, rotated rx 146.14 ry 0 rz 180 deg; joints [-11.684, -63.028, 110.007, 164.206, 48.077, -113.155]
  MoveL 3101 to (0, -37.84, 55.62) mm, rotated rx 143.54 ry 0 rz 180 deg; joints [-11.359, -63.724, 109.823, 164.421, 47.169, -115.728]
  MoveL 3102 to (-200, -37.84, 55.62) mm, rotated rx 143.54 ry 0 rz 180 deg; joints [-13.234, -74.551, 125.679, 163.192, 52.344, -116.005]
  MoveL 3103 to (-200, -38.32, 55.25) mm, rotated rx 140.94 ry 0 rz 180 deg; joints [-12.828, -75.369, 125.466, 163.468, 51.283, -118.547]
  MoveL 3104 to (0, -38.32, 55.25) mm, rotated rx 140.94 ry 0 rz 180 deg; joints [-11.007, -64.397, 109.636, 164.68, 46.275, -118.343]
  MoveL 3105 to (0, -38.78, 54.86) mm, rotated rx 138.33 ry 0 rz 180 deg; joints [-10.627, -65.047, 109.448, 164.988, 45.395, -121.005]
  MoveL 3106 to (-200, -38.78, 54.86) mm, rotated rx 138.33 ry 0 rz 180 deg; joints [-12.389, -76.158, 125.252, 163.794, 50.24, -121.14]
  MoveL 3107 to (-200, -39.22, 54.45) mm, rotated rx 135.73 ry 0 rz 180 deg; joints [-11.919, -76.916, 125.037, 164.172, 49.219, -123.783]
  MoveL 3108 to (0, -39.22, 54.45) mm, rotated rx 135.73 ry 0 rz 180 deg; joints [-10.221, -65.672, 109.259, 165.344, 44.534, -123.714]
  MoveL 3109 to (0, -39.63, 54.02) mm, rotated rx 133.12 ry 0 rz 180 deg; joints [-9.789, -66.271, 109.07, 165.751, 43.693, -126.473]
  MoveL 3110 to (-200, -39.63, 54.02) mm, rotated rx 133.12 ry 0 rz 180 deg; joints [-11.419, -77.642, 124.822, 164.604, 48.222, -126.482]
  MoveL 3111 to (-200, -40.03, 53.58) mm, rotated rx 130.52 ry 0 rz 180 deg; joints [-10.89, -78.334, 124.608, 165.093, 47.252, -129.24]
  MoveL 3112 to (0, -40.03, 53.58) mm, rotated rx 130.52 ry 0 rz 180 deg; joints [-9.332, -66.843, 108.882, 166.212, 42.874, -129.287]
  MoveL 3113 to (0, -40.41, 53.11) mm, rotated rx 127.91 ry 0 rz 180 deg; joints [-8.851, -67.387, 108.696, 166.726, 42.08, -132.156]
  MoveL 3114 to (-200, -40.41, 53.11) mm, rotated rx 127.91 ry 0 rz 180 deg; joints [-10.332, -78.993, 124.396, 165.64, 46.312, -132.059]
  MoveL 3115 to (-200, -40.77, 52.63) mm, rotated rx 125.31 ry 0 rz 180 deg; joints [-9.746, -79.616, 124.187, 166.248, 45.404, -134.941]
  MoveL 3116 to (0, -40.77, 52.63) mm, rotated rx 125.31 ry 0 rz 180 deg; joints [-8.347, -67.903, 108.512, 167.297, 41.312, -135.082]
  MoveL 3117 to (0, -41.11, 52.13) mm, rotated rx 122.7 ry 0 rz 180 deg; joints [-7.82, -68.389, 108.331, 167.926, 40.575, -138.068]
  MoveL 3118 to (-200, -41.11, 52.13) mm, rotated rx 122.7 ry 0 rz 180 deg; joints [-9.133, -80.203, 123.982, 166.919, 44.532, -137.891]
  MoveL 3119 to (-200, -41.42, 51.62) mm, rotated rx 120.1 ry 0 rz 180 deg; joints [-8.495, -80.753, 123.781, 167.653, 43.697, -140.907]
  MoveL 3120 to (0, -41.42, 51.62) mm, rotated rx 120.1 ry 0 rz 180 deg; joints [-7.271, -68.844, 108.155, 168.613, 39.87, -141.113]
  MoveL 3121 to (0, -41.71, 51.09) mm, rotated rx 117.5 ry 0 rz 180 deg; joints [-6.702, -69.269, 107.983, 169.358, 39.199, -144.219]
  MoveL 3122 to (-200, -41.71, 51.09) mm, rotated rx 117.5 ry 0 rz 180 deg; joints [-7.833, -81.265, 123.587, 168.452, 42.905, -143.992]
  MoveL 3123 to (-200, -41.97, 50.56) mm, rotated rx 114.89 ry 0 rz 180 deg; joints [-7.148, -81.739, 123.398, 169.316, 42.157, -147.147]
  MoveL 3124 to (0, -41.97, 50.56) mm, rotated rx 114.89 ry 0 rz 180 deg; joints [-6.114, -69.662, 107.816, 170.163, 38.566, -147.388]
  MoveL 3125 to (0, -42.21, 50.01) mm, rotated rx 112.29 ry 0 rz 180 deg; joints [-5.508, -70.023, 107.655, 171.025, 37.974, -150.616]
  MoveL 3126 to (-200, -42.21, 50.01) mm, rotated rx 112.29 ry 0 rz 180 deg; joints [-6.441, -82.174, 123.217, 170.245, 41.457, -150.371]
  MoveL 3127 to (-200, -42.43, 49.45) mm, rotated rx 109.68 ry 0 rz 180 deg; joints [-5.714, -82.569, 123.045, 171.237, 40.808, -153.663]
  MoveL 3128 to (0, -42.43, 49.45) mm, rotated rx 109.68 ry 0 rz 180 deg; joints [-4.885, -70.352, 107.502, 171.944, 37.424, -153.905]
  MoveL 3129 to (0, -42.62, 48.88) mm, rotated rx 107.08 ry 0 rz 180 deg; joints [-4.247, -70.647, 107.356, 172.917, 36.92, -157.249]
  MoveL 3130 to (-200, -42.62, 48.88) mm, rotated rx 107.08 ry 0 rz 180 deg; joints [-4.969, -82.924, 122.881, 172.29, 40.213, -157.02]
  MoveL 3131 to (-200, -42.78, 48.3) mm, rotated rx 104.47 ry 0 rz 180 deg; joints [-4.207, -83.238, 122.727, 173.402, 39.676, -160.438]
  MoveL 3132 to (0, -42.78, 48.3) mm, rotated rx 104.47 ry 0 rz 180 deg; joints [-3.596, -70.908, 107.218, 173.943, 36.463, -160.648]
  MoveL 3133 to (0, -42.92, 47.72) mm, rotated rx 101.87 ry 0 rz 180 deg; joints [-2.931, -71.135, 107.088, 175.016, 36.056, -164.099]
  MoveL 3134 to (-200, -42.92, 47.72) mm, rotated rx 101.87 ry 0 rz 180 deg; joints [-3.43, -83.511, 122.583, 174.568, 39.198, -163.917]
  MoveL 3135 to (-200, -43.03, 47.12) mm, rotated rx 99.27 ry 0 rz 180 deg; joints [-2.64, -83.743, 122.45, 175.783, 38.783, -167.446]
  MoveL 3136 to (0, -43.03, 47.12) mm, rotated rx 99.27 ry 0 rz 180 deg; joints [-2.255, -71.328, 106.968, 176.133, 35.701, -167.593]
  MoveL 3137 to (0, -43.11, 46.53) mm, rotated rx 96.66 ry 0 rz 180 deg; joints [-1.57, -71.487, 106.858, 177.288, 35.401, -171.128]
  MoveL 3138 to (-200, -43.11, 46.53) mm, rotated rx 96.66 ry 0 rz 180 deg; joints [-1.838, -83.933, 122.329, 177.042, 38.433, -171.021]
  MoveL 3139 to (-200, -43.17, 45.93) mm, rotated rx 94.06 ry 0 rz 180 deg; joints [-1.027, -84.081, 122.219, 178.337, 38.15, -174.636]
  MoveL 3140 to (0, -43.17, 45.93) mm, rotated rx 94.06 ry 0 rz 180 deg; joints [-0.877, -71.611, 106.757, 178.476, 35.156, -174.698]
  MoveL 3141 to (0, -43.2, 45.33) mm, rotated rx 91.45 ry 0 rz 180 deg; joints [-0.178, -71.7, 106.667, 179.689, 34.968, -178.293]
  MoveL 3142 to (-200, -43.2, 45.33) mm, rotated rx 91.45 ry 0 rz 180 deg; joints [-0.209, -84.187, 122.122, 179.66, 37.935, -178.28]
  MoveL 3143 to (-200, -43.2, 44.73) mm, rotated rx 90 ry 0 rz 180 deg; joints [0.263, -84.228, 122.073, -179.571, 37.846, 179.662]
  MoveL 3144 to (0, -43.2, 44.73) mm, rotated rx 90 ry 0 rz 180 deg; joints [0.225, -71.734, 106.622, -179.607, 34.888, 179.678]
  MoveL 3145 to (0, -43.2, 44.13) mm, rotated rx 90 ry 0 rz 180 deg; joints [0.25, -71.734, 106.622, -179.564, 34.888, 179.642]
  MoveL 3146 to (-200, -43.2, 44.13) mm, rotated rx 90 ry 0 rz 180 deg; joints [0.292, -84.228, 122.073, -179.524, 37.846, 179.624]
  MoveL 3147 to (-200, -43.2, 43.53) mm, rotated rx 90 ry 0 rz 180 deg; joints [0.322, -84.228, 122.073, -179.476, 37.846, 179.586]
  MoveL 3148 to (0, -43.2, 43.53) mm, rotated rx 90 ry 0 rz 180 deg; joints [0.275, -71.734, 106.622, -179.52, 34.888, 179.606]
  MoveL 3149 to (0, -43.2, 42.94) mm, rotated rx 90 ry 0 rz 180 deg; joints [0.3, -71.734, 106.621, -179.476, 34.888, 179.57]
  MoveL 3150 to (-200, -43.2, 42.94) mm, rotated rx 90 ry 0 rz 180 deg; joints [0.351, -84.228, 122.073, -179.428, 37.846, 179.548]
  MoveL 3151 to (-200, -43.2, 42.34) mm, rotated rx 90 ry 0 rz 180 deg; joints [0.38, -84.227, 122.073, -179.38, 37.847, 179.511]
  MoveL 3152 to (0, -43.2, 42.34) mm, rotated rx 90 ry 0 rz 180 deg; joints [0.325, -71.734, 106.621, -179.432, 34.889, 179.534]
  MoveL 3153 to (0, -43.2, 41.73) mm, rotated rx 90 ry 0 rz 180 deg; joints [0.35, -71.734, 106.621, -179.388, 34.889, 179.498]
  MoveL 3154 to (-200, -43.2, 41.73) mm, rotated rx 90 ry 0 rz 180 deg; joints [0.41, -84.227, 122.072, -179.332, 37.847, 179.473]
  MoveL 3155 to (-200, -43.2, 41.13) mm, rotated rx 90 ry 0 rz 180 deg; joints [0.439, -84.227, 122.072, -179.285, 37.847, 179.435]
  MoveL 3156 to (0, -43.2, 41.13) mm, rotated rx 90 ry 0 rz 180 deg; joints [0.375, -71.733, 106.62, -179.344, 34.889, 179.462]
  MoveL 3157 to (0, -43.2, 40.53) mm, rotated rx 90 ry 0 rz 180 deg; joints [0.4, -71.733, 106.62, -179.301, 34.889, 179.426]
  MoveL 3158 to (-200, -43.2, 40.53) mm, rotated rx 90 ry 0 rz 180 deg; joints [0.468, -84.227, 122.072, -179.237, 37.847, 179.397]
  MoveL 3159 to (-200, -43.2, 39.94) mm, rotated rx 90 ry 0 rz 180 deg; joints [0.498, -84.226, 122.071, -179.189, 37.848, 179.36]
  MoveL 3160 to (0, -43.2, 39.94) mm, rotated rx 90 ry 0 rz 180 deg; joints [0.425, -71.733, 106.62, -179.257, 34.889, 179.39]
  MoveL 3161 to (0, -43.2, 39.34) mm, rotated rx 90 ry 0 rz 180 deg; joints [0.45, -71.732, 106.619, -179.213, 34.889, 179.355]
  MoveL 3162 to (-200, -43.2, 39.34) mm, rotated rx 90 ry 0 rz 180 deg; joints [0.527, -84.226, 122.071, -179.141, 37.848, 179.322]
  MoveL 3163 to (-200, -43.2, 38.73) mm, rotated rx 90 ry 0 rz 180 deg; joints [0.556, -84.226, 122.07, -179.093, 37.848, 179.284]
  MoveL 3164 to (0, -43.2, 38.73) mm, rotated rx 90 ry 0 rz 180 deg; joints [0.475, -71.732, 106.619, -179.169, 34.89, 179.319]
  MoveL 3165 to (0, -43.2, 38.13) mm, rotated rx 90 ry 0 rz 180 deg; joints [0.5, -71.732, 106.618, -179.125, 34.89, 179.283]
  MoveL 3166 to (-200, -43.2, 38.13) mm, rotated rx 90 ry 0 rz 180 deg; joints [0.586, -84.225, 122.07, -179.046, 37.849, 179.246]
  MoveL 3167 to (-200, -43.2, 37.53) mm, rotated rx 90 ry 0 rz 180 deg; joints [0.615, -84.225, 122.07, -178.998, 37.849, 179.209]
  MoveL 3168 to (0, -43.2, 37.53) mm, rotated rx 90 ry 0 rz 180 deg; joints [0.525, -71.732, 106.618, -179.082, 34.89, 179.247]
  MoveL 3169 to (0, -43.2, 36.94) mm, rotated rx 90 ry 0 rz 180 deg; joints [0.55, -71.731, 106.618, -179.038, 34.89, 179.211]
  MoveL 3170 to (-200, -43.2, 36.94) mm, rotated rx 90 ry 0 rz 180 deg; joints [0.644, -84.224, 122.069, -178.95, 37.849, 179.171]
  MoveL 3171 to (-200, -43.2, 36.34) mm, rotated rx 90 ry 0 rz 180 deg; joints [0.674, -84.224, 122.069, -178.902, 37.85, 179.133]
  MoveL 3172 to (0, -43.2, 36.34) mm, rotated rx 90 ry 0 rz 180 deg; joints [0.575, -71.731, 106.617, -178.994, 34.89, 179.175]
  MoveL 3173 to (0, -43.2, 35.73) mm, rotated rx 90 ry 0 rz 180 deg; joints [0.6, -71.73, 106.617, -178.95, 34.891, 179.139]
  MoveL 3174 to (-200, -43.2, 35.73) mm, rotated rx 90 ry 0 rz 180 deg; joints [0.703, -84.223, 122.068, -178.854, 37.85, 179.095]
  MoveL 3175 to (-200, -43.2, 35.13) mm, rotated rx 90 ry 0 rz 180 deg; joints [0.732, -84.223, 122.068, -178.807, 37.851, 179.058]
  MoveL 3176 to (0, -43.2, 35.13) mm, rotated rx 90 ry 0 rz 180 deg; joints [0.625, -71.73, 106.616, -178.906, 34.891, 179.103]
  MoveL 3177 to (0, -43.2, 34.53) mm, rotated rx 90 ry 0 rz 180 deg; joints [0.651, -71.73, 106.615, -178.863, 34.891, 179.067]
  MoveL 3178 to (-200, -43.2, 34.53) mm, rotated rx 90 ry 0 rz 180 deg; joints [0.762, -84.222, 122.067, -178.759, 37.851, 179.02]
  MoveL 3179 to (-200, -43.2, 33.94) mm, rotated rx 90 ry 0 rz 180 deg; joints [0.791, -84.222, 122.066, -178.711, 37.851, 178.982]
  MoveL 3180 to (0, -43.2, 33.94) mm, rotated rx 90 ry 0 rz 180 deg; joints [0.676, -71.729, 106.615, -178.819, 34.891, 179.031]
  MoveL 3181 to (0, -43.2, 33.34) mm, rotated rx 90 ry 0 rz 180 deg; joints [0.701, -71.729, 106.614, -178.775, 34.892, 178.995]
  MoveL 3182 to (-200, -43.2, 33.34) mm, rotated rx 90 ry 0 rz 180 deg; joints [0.82, -84.221, 122.066, -178.663, 37.852, 178.944]
  MoveL 3183 to (-200, -43.2, 32.73) mm, rotated rx 90 ry 0 rz 180 deg; joints [0.85, -84.221, 122.065, -178.615, 37.852, 178.907]
  MoveL 3184 to (0, -43.2, 32.73) mm, rotated rx 90 ry 0 rz 180 deg; joints [0.726, -71.728, 106.614, -178.731, 34.892, 178.959]
  MoveL 3185 to (0, -43.2, 32.13) mm, rotated rx 90 ry 0 rz 180 deg; joints [0.751, -71.728, 106.613, -178.687, 34.892, 178.923]
  MoveL 3186 to (-200, -43.2, 32.13) mm, rotated rx 90 ry 0 rz 180 deg; joints [0.879, -84.22, 122.064, -178.568, 37.853, 178.869]
  MoveL 3187 to (-200, -43.2, 31.54) mm, rotated rx 90 ry 0 rz 180 deg; joints [0.908, -84.22, 122.064, -178.52, 37.853, 178.831]
  MoveL 3188 to (0, -43.2, 31.54) mm, rotated rx 90 ry 0 rz 180 deg; joints [0.776, -71.727, 106.612, -178.644, 34.893, 178.887]
  MoveL 3189 to (0, -43.2, 30.93) mm, rotated rx 90 ry 0 rz 180 deg; joints [0.801, -71.727, 106.612, -178.6, 34.893, 178.852]
  MoveL 3190 to (-200, -43.2, 30.93) mm, rotated rx 90 ry 0 rz 180 deg; joints [0.938, -84.219, 122.063, -178.472, 37.854, 178.794]
  MoveL 3191 to (-200, -43.2, 30.34) mm, rotated rx 90 ry 0 rz 180 deg; joints [0.967, -84.218, 122.062, -178.424, 37.855, 178.756]
  MoveL 3192 to (0, -43.2, 30.34) mm, rotated rx 90 ry 0 rz 180 deg; joints [0.826, -71.726, 106.611, -178.556, 34.893, 178.816]
  MoveL 3193 to (0, -43.2, 29.73) mm, rotated rx 90 ry 0 rz 180 deg; joints [0.851, -71.726, 106.61, -178.512, 34.894, 178.78]
  MoveL 3194 to (-200, -43.2, 29.73) mm, rotated rx 90 ry 0 rz 180 deg; joints [0.996, -84.218, 122.062, -178.377, 37.855, 178.718]
  MoveL 3195 to (-200, -43.2, 29.14) mm, rotated rx 90 ry 0 rz 180 deg; joints [1.025, -84.217, 122.061, -178.329, 37.856, 178.68]
  MoveL 3196 to (0, -43.2, 29.14) mm, rotated rx 90 ry 0 rz 180 deg; joints [0.876, -71.725, 106.609, -178.469, 34.894, 178.744]
  MoveL 3197 to (0, -43.2, 28.54) mm, rotated rx 90 ry 0 rz 180 deg; joints [0.901, -71.725, 106.609, -178.425, 34.894, 178.708]
  MoveL 3198 to (-200, -43.2, 28.54) mm, rotated rx 90 ry 0 rz 180 deg; joints [1.055, -84.216, 122.06, -178.281, 37.856, 178.643]
  MoveL 3199 to (-200, -43.2, 27.93) mm, rotated rx 90 ry 0 rz 180 deg; joints [1.084, -84.216, 122.059, -178.233, 37.857, 178.605]
  MoveL 3200 to (0, -43.2, 27.93) mm, rotated rx 90 ry 0 rz 180 deg; joints [0.926, -71.724, 106.608, -178.381, 34.895, 178.672]
  MoveL 3201 to (0, -43.2, 27.34) mm, rotated rx 90 ry 0 rz 180 deg; joints [0.951, -71.723, 106.607, -178.337, 34.895, 178.636]
  MoveL 3202 to (-200, -43.2, 27.34) mm, rotated rx 90 ry 0 rz 180 deg; joints [1.113, -84.215, 122.058, -178.185, 37.858, 178.567]
  MoveL 3203 to (-200, -43.2, 26.73) mm, rotated rx 90 ry 0 rz 180 deg; joints [1.143, -84.214, 122.058, -178.138, 37.858, 178.529]
  MoveL 3204 to (0, -43.2, 26.73) mm, rotated rx 90 ry 0 rz 180 deg; joints [0.976, -71.723, 106.606, -178.293, 34.895, 178.6]
  MoveL 3205 to (0, -43.2, 26.14) mm, rotated rx 90 ry 0 rz 180 deg; joints [1.001, -71.722, 106.605, -178.25, 34.896, 178.564]
  MoveL 3206 to (-200, -43.2, 26.14) mm, rotated rx 90 ry 0 rz 180 deg; joints [1.172, -84.213, 122.057, -178.09, 37.859, 178.492]
  MoveL 3207 to (-200, -43.2, 25.54) mm, rotated rx 90 ry 0 rz 180 deg; joints [1.201, -84.213, 122.056, -178.042, 37.86, 178.454]
  MoveL 3208 to (0, -43.2, 25.54) mm, rotated rx 90 ry 0 rz 180 deg; joints [1.026, -71.722, 106.604, -178.206, 34.896, 178.528]
  MoveL 3209 to (0, -43.2, 24.93) mm, rotated rx 90 ry 0 rz 180 deg; joints [1.051, -71.721, 106.604, -178.162, 34.897, 178.492]
  MoveL 3210 to (-200, -43.2, 24.93) mm, rotated rx 90 ry 0 rz 180 deg; joints [1.231, -84.212, 122.055, -177.994, 37.86, 178.416]
  MoveL 3211 to (-200, -43.2, 24.34) mm, rotated rx 90 ry 0 rz 180 deg; joints [1.26, -84.211, 122.054, -177.947, 37.861, 178.379]
  MoveL 3212 to (0, -43.2, 24.34) mm, rotated rx 90 ry 0 rz 180 deg; joints [1.076, -71.72, 106.603, -178.118, 34.897, 178.456]
  MoveL 3213 to (0, -43.2, 23.73) mm, rotated rx 90 ry 0 rz 180 deg; joints [1.101, -71.719, 106.602, -178.074, 34.897, 178.421]
  MoveL 3214 to (-200, -43.2, 23.73) mm, rotated rx 90 ry 0 rz 180 deg; joints [1.289, -84.21, 122.053, -177.899, 37.862, 178.341]
  MoveL 3215 to (-200, -43.2, 23.14) mm, rotated rx 90 ry 0 rz 180 deg; joints [1.319, -84.209, 122.052, -177.851, 37.862, 178.303]
  MoveL 3216 to (0, -43.2, 23.14) mm, rotated rx 90 ry 0 rz 180 deg; joints [1.127, -71.719, 106.601, -178.031, 34.898, 178.385]
  MoveL 3217 to (0, -43.2, 22.54) mm, rotated rx 90 ry 0 rz 180 deg; joints [1.152, -71.718, 106.6, -177.987, 34.898, 178.349]
  MoveL 3218 to (-200, -43.2, 22.54) mm, rotated rx 90 ry 0 rz 180 deg; joints [1.348, -84.208, 122.051, -177.803, 37.863, 178.266]
  MoveL 3219 to (-200, -43.2, 21.93) mm, rotated rx 90 ry 0 rz 180 deg; joints [1.377, -84.207, 122.05, -177.756, 37.864, 178.228]
  MoveL 3220 to (0, -43.2, 21.93) mm, rotated rx 90 ry 0 rz 180 deg; joints [1.177, -71.717, 106.599, -177.943, 34.899, 178.313]
  MoveL 3221 to (0, -43.2, 21.34) mm, rotated rx 90 ry 0 rz 180 deg; joints [1.202, -71.717, 106.598, -177.899, 34.899, 178.277]
  MoveL 3222 to (-200, -43.2, 21.34) mm, rotated rx 90 ry 0 rz 180 deg; joints [1.407, -84.206, 122.049, -177.708, 37.865, 178.19]
  MoveL 3223 to (-200, -43.2, 20.73) mm, rotated rx 90 ry 0 rz 180 deg; joints [1.436, -84.205, 122.048, -177.66, 37.866, 178.152]
  MoveL 3224 to (0, -43.2, 20.73) mm, rotated rx 90 ry 0 rz 180 deg; joints [1.227, -71.716, 106.597, -177.856, 34.9, 178.241]
  MoveL 3225 to (0, -43.2, 20.14) mm, rotated rx 90 ry 0 rz 180 deg; joints [1.252, -71.715, 106.596, -177.812, 34.9, 178.205]
  MoveL 3226 to (-200, -43.2, 20.14) mm, rotated rx 90 ry 0 rz 180 deg; joints [1.465, -84.204, 122.047, -177.612, 37.866, 178.115]
  MoveL 3227 to (-200, -43.2, 19.54) mm, rotated rx 90 ry 0 rz 180 deg; joints [1.495, -84.203, 122.046, -177.565, 37.867, 178.077]
  MoveL 3228 to (0, -43.2, 19.54) mm, rotated rx 90 ry 0 rz 180 deg; joints [1.277, -71.714, 106.594, -177.768, 34.901, 178.169]
  MoveL 3229 to (0, -43.2, 18.93) mm, rotated rx 90 ry 0 rz 180 deg; joints [1.302, -71.713, 106.593, -177.724, 34.901, 178.133]
  MoveL 3230 to (-200, -43.2, 18.93) mm, rotated rx 90 ry 0 rz 180 deg; joints [1.524, -84.202, 122.045, -177.517, 37.868, 178.039]
  MoveL 3231 to (-200, -43.2, 18.34) mm, rotated rx 90 ry 0 rz 180 deg; joints [1.553, -84.201, 122.043, -177.469, 37.869, 178.002]
  MoveL 3232 to (0, -43.2, 18.34) mm, rotated rx 90 ry 0 rz 180 deg; joints [1.327, -71.712, 106.592, -177.681, 34.902, 178.097]
  MoveL 3233 to (0, -43.2, 17.73) mm, rotated rx 90 ry 0 rz 180 deg; joints [1.352, -71.712, 106.591, -177.637, 34.902, 178.062]
  MoveL 3234 to (-200, -43.2, 17.73) mm, rotated rx 90 ry 0 rz 180 deg; joints [1.583, -84.2, 122.042, -177.422, 37.87, 177.964]
  MoveL 3235 to (-200, -43.2, 17.14) mm, rotated rx 90 ry 0 rz 180 deg; joints [1.612, -84.199, 122.041, -177.374, 37.871, 177.926]
  MoveL 3236 to (0, -43.2, 17.14) mm, rotated rx 90 ry 0 rz 180 deg; joints [1.377, -71.711, 106.59, -177.593, 34.903, 178.026]
  MoveL 3237 to (0, -43.2, 16.54) mm, rotated rx 90 ry 0 rz 180 deg; joints [1.402, -71.71, 106.589, -177.549, 34.903, 177.99]
  MoveL 3238 to (-200, -43.2, 16.54) mm, rotated rx 90 ry 0 rz 180 deg; joints [1.641, -84.198, 122.04, -177.326, 37.872, 177.889]
  MoveL 3239 to (-200, -43.2, 15.94) mm, rotated rx 90 ry 0 rz 180 deg; joints [1.67, -84.197, 122.039, -177.278, 37.873, 177.851]
  MoveL 3240 to (0, -43.2, 15.94) mm, rotated rx 90 ry 0 rz 180 deg; joints [1.427, -71.709, 106.587, -177.506, 34.904, 177.954]
  MoveL 3241 to (0, -43.2, 15.34) mm, rotated rx 90 ry 0 rz 180 deg; joints [1.452, -71.708, 106.586, -177.462, 34.905, 177.918]
  MoveL 3242 to (-200, -43.2, 15.34) mm, rotated rx 90 ry 0 rz 180 deg; joints [1.7, -84.196, 122.037, -177.231, 37.874, 177.813]
  MoveL 3243 to (-200, -43.2, 14.73) mm, rotated rx 88.85 ry 0 rz 180 deg; joints [2.081, -84.206, 121.987, -176.606, 37.83, 176.166]
  MoveL 3244 to (0, -43.2, 14.73) mm, rotated rx 88.85 ry 0 rz 180 deg; joints [1.778, -71.717, 106.538, -176.889, 34.861, 176.295]
  MoveL 3245 to (0, -43.17, 14.13) mm, rotated rx 86.24 ry 0 rz 180 deg; joints [2.484, -71.713, 106.439, -175.646, 34.804, 172.666]
  MoveL 3246 to (-200, -43.17, 14.13) mm, rotated rx 86.24 ry 0 rz 180 deg; joints [2.907, -84.201, 121.885, -175.252, 37.779, 172.487]
  MoveL 3247 to (-200, -43.12, 13.54) mm, rotated rx 83.64 ry 0 rz 180 deg; joints [3.733, -84.153, 121.795, -173.902, 37.799, 168.814]
  MoveL 3248 to (0, -43.12, 13.54) mm, rotated rx 83.64 ry 0 rz 180 deg; joints [3.19, -71.675, 106.352, -174.405, 34.805, 169.04]
  MoveL 3249 to (0, -43.04, 12.94) mm, rotated rx 81.03 ry 0 rz 180 deg; joints [3.896, -71.602, 106.276, -173.174, 34.865, 165.425]
  MoveL 3250 to (-200, -43.04, 12.94) mm, rotated rx 81.03 ry 0 rz 180 deg; joints [4.558, -84.064, 121.719, -172.565, 37.889, 165.155]
  MoveL 3251 to (-200, -42.93, 12.35) mm, rotated rx 78.43 ry 0 rz 180 deg; joints [5.38, -83.934, 121.656, -171.249, 38.047, 161.518]
  MoveL 3252 to (0, -42.93, 12.35) mm, rotated rx 78.43 ry 0 rz 180 deg; joints [4.599, -71.494, 106.211, -171.96, 34.982, 161.828]
  MoveL 3253 to (0, -42.8, 11.77) mm, rotated rx 75.83 ry 0 rz 180 deg; joints [5.299, -71.352, 106.158, -170.771, 35.156, 158.259]
  MoveL 3254 to (-200, -42.8, 11.77) mm, rotated rx 75.83 ry 0 rz 180 deg; joints [6.196, -83.763, 121.607, -169.965, 38.273, 157.917]
  MoveL 3255 to (-200, -42.64, 11.19) mm, rotated rx 73.22 ry 0 rz 180 deg; joints [7.005, -83.551, 121.571, -168.718, 38.564, 154.356]
  MoveL 3256 to (0, -42.64, 11.19) mm, rotated rx 73.22 ry 0 rz 180 deg; joints [5.992, -71.177, 106.116, -169.614, 35.385, 154.724]
  MoveL 3257 to (0, -42.45, 10.62) mm, rotated rx 70.62 ry 0 rz 180 deg; joints [6.678, -70.968, 106.086, -168.495, 35.667, 151.228]
  MoveL 3258 to (-200, -42.45, 10.62) mm, rotated rx 70.62 ry 0 rz 180 deg; joints [7.805, -83.299, 121.548, -167.515, 38.917, 150.843]
  MoveL 3259 to (-200, -42.24, 10.06) mm, rotated rx 68.01 ry 0 rz 180 deg; joints [8.593, -83.008, 121.538, -166.364, 39.331, 147.385]
  MoveL 3260 to (0, -42.24, 10.06) mm, rotated rx 68.01 ry 0 rz 180 deg; joints [7.356, -70.725, 106.067, -167.42, 36.001, 147.779]
  MoveL 3261 to (0, -42, 9.51) mm, rotated rx 65.41 ry 0 rz 180 deg; joints [8.023, -70.451, 106.06, -166.392, 36.385, 144.381]
  MoveL 3262 to (-200, -42, 9.51) mm, rotated rx 65.41 ry 0 rz 180 deg; joints [9.369, -82.677, 121.541, -165.268, 39.803, 143.987]
  MoveL 3263 to (-200, -41.74, 8.97) mm, rotated rx 62.8 ry 0 rz 180 deg; joints [10.13, -82.309, 121.557, -164.231, 40.329, 140.655]
  MoveL 3264 to (0, -41.74, 8.97) mm, rotated rx 62.8 ry 0 rz 180 deg; joints [8.677, -70.144, 106.063, -165.417, 36.815, 141.039]
  MoveL 3265 to (0, -41.45, 8.44) mm, rotated rx 60.2 ry 0 rz 180 deg; joints [9.319, -69.806, 106.077, -164.497, 37.29, 137.756]
  MoveL 3266 to (-200, -41.45, 8.44) mm, rotated rx 60.2 ry 0 rz 180 deg; joints [10.874, -81.903, 121.584, -163.256, 40.906, 137.39]
  MoveL 3267 to (-200, -41.15, 7.93) mm, rotated rx 57.6 ry 0 rz 180 deg; joints [11.601, -81.46, 121.623, -162.345, 41.531, 134.193]
  MoveL 3268 to (0, -41.15, 7.93) mm, rotated rx 57.6 ry 0 rz 180 deg; joints [9.946, -69.437, 106.102, -163.634, 37.806, 134.532]
  MoveL 3269 to (0, -40.81, 7.43) mm, rotated rx 54.99 ry 0 rz 180 deg; joints [10.557, -69.038, 106.136, -162.83, 38.362, 131.372]
  MoveL 3270 to (-200, -40.81, 7.43) mm, rotated rx 54.99 ry 0 rz 180 deg; joints [12.308, -80.981, 121.674, -161.498, 42.201, 131.069]
  MoveL 3271 to (-200, -40.46, 6.94) mm, rotated rx 52.39 ry 0 rz 180 deg; joints [12.994, -80.466, 121.735, -160.717, 42.913, 128.015]
  MoveL 3272 to (0, -40.46, 6.94) mm, rotated rx 52.39 ry 0 rz 180 deg; joints [11.151, -68.609, 106.18, -162.085, 38.955, 128.275]
  MoveL 3273 to (0, -40.08, 6.48) mm, rotated rx 49.78 ry 0 rz 180 deg; joints [11.727, -68.152, 106.233, -161.399, 39.583, 125.241]
  MoveL 3274 to (-200, -40.08, 6.48) mm, rotated rx 49.78 ry 0 rz 180 deg; joints [13.658, -79.918, 121.806, -160.001, 43.664, 125.032]
  MoveL 3275 to (-200, -39.68, 6.03) mm, rotated rx 47.18 ry 0 rz 180 deg; joints [14.299, -79.336, 121.886, -159.348, 44.45, 122.118]
  MoveL 3276 to (0, -39.68, 6.03) mm, rotated rx 47.18 ry 0 rz 180 deg; joints [12.283, -67.667, 106.295, -160.773, 40.241, 122.27]
  MoveL 3277 to (0, -39.26, 5.6) mm, rotated rx 44.57 ry 0 rz 180 deg; joints [12.819, -67.155, 106.365, -160.204, 40.929, 119.361]
  MoveL 3278 to (-200, -39.26, 5.6) mm, rotated rx 44.57 ry 0 rz 180 deg; joints [14.916, -78.722, 121.976, -158.757, 45.269, 119.273]
  MoveL 3279 to (-200, -38.83, 5.19) mm, rotated rx 41.97 ry 0 rz 180 deg; joints [15.507, -78.075, 122.073, -158.227, 46.117, 116.493]
  MoveL 3280 to (0, -38.83, 5.19) mm, rotated rx 41.97 ry 0 rz 180 deg; joints [13.333, -66.617, 106.443, -159.693, 41.644, 116.511]
  MoveL 3281 to (0, -38.37, 4.79) mm, rotated rx 39.37 ry 0 rz 180 deg; joints [13.826, -66.053, 106.528, -159.237, 42.383, 113.72]
  MoveL 3282 to (-200, -38.37, 4.79) mm, rotated rx 39.37 ry 0 rz 180 deg; joints [16.071, -77.399, 122.178, -157.755, 46.993, 113.777]
  MoveL 3283 to (-200, -37.9, 4.42) mm, rotated rx 36.76 ry 0 rz 180 deg; joints [16.609, -76.694, 122.29, -157.339, 47.893, 111.122]
  MoveL 3284 to (0, -37.9, 4.42) mm, rotated rx 36.76 ry 0 rz 180 deg; joints [14.295, -65.465, 106.619, -158.834, 43.144, 110.986]
  MoveL 3285 to (0, -37.41, 4.08) mm, rotated rx 34.16 ry 0 rz 180 deg; joints [14.74, -64.854, 106.716, -158.484, 43.925, 108.304]
  MoveL 3286 to (-200, -37.41, 4.08) mm, rotated rx 34.16 ry 0 rz 180 deg; joints [17.118, -75.96, 122.408, -156.976, 48.816, 108.523]
  MoveL 3287 to (-200, -36.91, 3.75) mm, rotated rx 31.55 ry 0 rz 180 deg; joints [17.599, -75.199, 122.532, -156.665, 49.758, 105.98]
  MoveL 3288 to (0, -36.91, 3.75) mm, rotated rx 31.55 ry 0 rz 180 deg; joints [15.161, -64.221, 106.819, -158.183, 44.725, 105.675]
  MoveL 3289 to (0, -36.39, 3.45) mm, rotated rx 28.95 ry 0 rz 180 deg; joints [15.557, -63.566, 106.926, -157.929, 45.54, 103.093]
  MoveL 3290 to (-200, -36.39, 3.45) mm, rotated rx 28.95 ry 0 rz 180 deg; joints [18.051, -74.412, 122.66, -156.402, 50.718, 103.487]
  MoveL 3291 to (-200, -35.86, 3.17) mm, rotated rx 26.34 ry 0 rz 180 deg; joints [18.472, -73.601, 122.793, -156.186, 51.694, 101.043]
  MoveL 3292 to (0, -35.86, 3.17) mm, rotated rx 26.34 ry 0 rz 180 deg; joints [15.926, -62.891, 107.038, -157.721, 46.369, 100.558]
  MoveL 3293 to (0, -35.31, 2.92) mm, rotated rx 23.74 ry 0 rz 180 deg; joints [16.27, -62.196, 107.153, -157.557, 47.211, 98.065]
  MoveL 3294 to (-200, -35.31, 2.92) mm, rotated rx 23.74 ry 0 rz 180 deg; joints [18.863, -72.767, 122.928, -156.013, 52.683, 98.643]
  MoveL 3295 to (-200, -34.76, 2.69) mm, rotated rx 21.13 ry 0 rz 180 deg; joints [19.224, -71.91, 123.067, -155.882, 53.685, 96.285]
  MoveL 3296 to (0, -34.76, 2.69) mm, rotated rx 21.13 ry 0 rz 180 deg; joints [16.587, -61.484, 107.271, -157.433, 48.063, 95.612]
  MoveL 3297 to (0, -34.2, 2.48) mm, rotated rx 18.53 ry 0 rz 180 deg; joints [16.877, -60.755, 107.392, -157.349, 48.925, 93.197]
  MoveL 3298 to (-200, -34.2, 2.48) mm, rotated rx 18.53 ry 0 rz 180 deg; joints [19.553, -71.033, 123.207, -155.79, 54.697, 93.965]
  MoveL 3299 to (-200, -33.62, 2.31) mm, rotated rx 15.93 ry 0 rz 180 deg; joints [19.85, -70.137, 123.349, -155.735, 55.718, 91.679]
  MoveL 3300 to (0, -33.62, 2.31) mm, rotated rx 15.93 ry 0 rz 180 deg; joints [17.139, -60.011, 107.515, -157.303, 49.794, 90.817]
  MoveL 3301 to (0, -33.04, 2.15) mm, rotated rx 13.32 ry 0 rz 180 deg; joints [17.373, -59.252, 107.639, -157.292, 50.669, 88.466]
  MoveL 3302 to (-200, -33.04, 2.15) mm, rotated rx 13.32 ry 0 rz 180 deg; joints [20.116, -69.222, 123.492, -155.716, 56.747, 89.425]
  MoveL 3303 to (-200, -32.45, 2.03) mm, rotated rx 10.72 ry 0 rz 180 deg; joints [20.35, -68.291, 123.635, -155.729, 57.78, 87.199]
  MoveL 3304 to (0, -32.45, 2.03) mm, rotated rx 10.72 ry 0 rz 180 deg; joints [17.58, -58.48, 107.764, -157.315, 51.549, 86.146]
  MoveL 3305 to (0, -31.86, 1.93) mm, rotated rx 8.11 ry 0 rz 180 deg; joints [17.758, -57.697, 107.89, -157.369, 52.432, 83.852]
  MoveL 3306 to (-200, -31.86, 1.93) mm, rotated rx 8.11 ry 0 rz 180 deg; joints [20.551, -67.346, 123.777, -155.775, 58.819, 84.999]
  MoveL 3307 to (-200, -31.27, 1.86) mm, rotated rx 5.51 ry 0 rz 180 deg; joints [20.72, -66.387, 123.919, -155.851, 59.861, 82.821]
  MoveL 3308 to (0, -31.27, 1.86) mm, rotated rx 5.51 ry 0 rz 180 deg; joints [17.907, -56.903, 108.015, -157.455, 53.317, 81.58]
  MoveL 3309 to (0, -30.67, 1.82) mm, rotated rx 2.9 ry 0 rz 180 deg; joints [18.028, -56.1, 108.14, -157.57, 54.203, 79.33]
  MoveL 3310 to (-200, -30.67, 1.82) mm, rotated rx 2.9 ry 0 rz 180 deg; joints [20.857, -65.417, 124.059, -155.955, 60.904, 80.663]
  MoveL 3311 to (-200, -30.07, 1.8) mm, rotated rx 0.3 ry 0 rz 180 deg; joints [20.961, -64.437, 124.198, -156.087, 61.948, 78.521]
  MoveL 3312 to (0, -30.07, 1.8) mm, rotated rx 0.3 ry 0 rz 180 deg; joints [18.12, -55.29, 108.265, -157.712, 55.089, 77.099]
  MoveL 3313 to (0, -29.47, 1.8) mm, rotated rx 0 ry 0 rz 180 deg; joints [18.129, -55.172, 108.285, -157.739, 55.219, 76.857]
  MoveL 3314 to (-200, -29.47, 1.8) mm, rotated rx 0 ry 0 rz 180 deg; joints [20.971, -64.293, 124.22, -156.112, 62.101, 78.292]
  MoveL 3315 to (-200, -28.87, 1.8) mm, rotated rx 0 ry 0 rz 180 deg; joints [20.971, -64.259, 124.227, -156.12, 62.138, 78.31]
  MoveL 3316 to (0, -28.87, 1.8) mm, rotated rx 0 ry 0 rz 180 deg; joints [18.129, -55.144, 108.291, -157.748, 55.251, 76.872]
  MoveL 3317 to (0, -28.27, 1.8) mm, rotated rx 0 ry 0 rz 180 deg; joints [18.129, -55.116, 108.297, -157.757, 55.282, 76.888]
  MoveL 3318 to (-200, -28.27, 1.8) mm, rotated rx 0 ry 0 rz 180 deg; joints [20.971, -64.225, 124.233, -156.129, 62.175, 78.329]
  MoveL 3319 to (-200, -27.67, 1.8) mm, rotated rx 0 ry 0 rz 180 deg; joints [20.971, -64.191, 124.24, -156.138, 62.213, 78.348]
  MoveL 3320 to (0, -27.67, 1.8) mm, rotated rx 0 ry 0 rz 180 deg; joints [18.129, -55.088, 108.304, -157.765, 55.314, 76.904]
  MoveL 3321 to (0, -27.07, 1.8) mm, rotated rx 0 ry 0 rz 180 deg; joints [18.129, -55.06, 108.31, -157.774, 55.346, 76.92]
  MoveL 3322 to (-200, -27.07, 1.8) mm, rotated rx 0 ry 0 rz 180 deg; joints [20.971, -64.157, 124.247, -156.146, 62.25, 78.366]
  MoveL 3323 to (-200, -26.47, 1.8) mm, rotated rx 0 ry 0 rz 180 deg; joints [20.971, -64.123, 124.254, -156.155, 62.287, 78.385]
  MoveL 3324 to (0, -26.47, 1.8) mm, rotated rx 0 ry 0 rz 180 deg; joints [18.129, -55.032, 108.316, -157.783, 55.377, 76.935]
  MoveL 3325 to (0, -25.87, 1.8) mm, rotated rx 0 ry 0 rz 180 deg; joints [18.129, -55.004, 108.322, -157.792, 55.409, 76.951]
  MoveL 3326 to (-200, -25.87, 1.8) mm, rotated rx 0 ry 0 rz 180 deg; joints [20.971, -64.089, 124.26, -156.164, 62.324, 78.404]
  MoveL 3327 to (-200, -25.27, 1.8) mm, rotated rx 0 ry 0 rz 180 deg; joints [20.971, -64.055, 124.267, -156.172, 62.362, 78.422]
  MoveL 3328 to (0, -25.27, 1.8) mm, rotated rx 0 ry 0 rz 180 deg; joints [18.129, -54.976, 108.328, -157.801, 55.441, 76.967]
  MoveL 3329 to (0, -24.67, 1.8) mm, rotated rx 0 ry 0 rz 180 deg; joints [18.129, -54.948, 108.334, -157.81, 55.472, 76.982]
  MoveL 3330 to (-200, -24.67, 1.8) mm, rotated rx 0 ry 0 rz 180 deg; joints [20.971, -64.021, 124.274, -156.181, 62.399, 78.441]
  MoveL 3331 to (-200, -24.07, 1.8) mm, rotated rx 0 ry 0 rz 180 deg; joints [20.971, -63.987, 124.28, -156.19, 62.436, 78.459]
  MoveL 3332 to (0, -24.07, 1.8) mm, rotated rx 0 ry 0 rz 180 deg; joints [18.129, -54.92, 108.341, -157.819, 55.504, 76.998]
  MoveL 3333 to (0, -23.47, 1.8) mm, rotated rx 0 ry 0 rz 180 deg; joints [18.129, -54.892, 108.347, -157.828, 55.535, 77.014]
  MoveL 3334 to (-200, -23.47, 1.8) mm, rotated rx 0 ry 0 rz 180 deg; joints [20.971, -63.953, 124.287, -156.198, 62.473, 78.478]
  MoveL 3335 to (-200, -22.87, 1.8) mm, rotated rx 0 ry 0 rz 180 deg; joints [20.971, -63.919, 124.293, -156.207, 62.51, 78.496]
  MoveL 3336 to (0, -22.87, 1.8) mm, rotated rx 0 ry 0 rz 180 deg; joints [18.129, -54.864, 108.353, -157.837, 55.567, 77.029]
  MoveL 3337 to (0, -22.27, 1.8) mm, rotated rx 0 ry 0 rz 180 deg; joints [18.129, -54.835, 108.359, -157.845, 55.599, 77.045]
  MoveL 3338 to (-200, -22.27, 1.8) mm, rotated rx 0 ry 0 rz 180 deg; joints [20.971, -63.885, 124.3, -156.215, 62.548, 78.515]
  MoveL 3339 to (-200, -21.67, 1.8) mm, rotated rx 0 ry 0 rz 180 deg; joints [20.971, -63.85, 124.306, -156.224, 62.585, 78.533]
  MoveL 3340 to (0, -21.67, 1.8) mm, rotated rx 0 ry 0 rz 180 deg; joints [18.129, -54.807, 108.365, -157.854, 55.63, 77.06]
  MoveL 3341 to (0, -21.07, 1.8) mm, rotated rx 0 ry 0 rz 180 deg; joints [18.129, -54.779, 108.37, -157.863, 55.662, 77.076]
  MoveL 3342 to (-200, -21.07, 1.8) mm, rotated rx 0 ry 0 rz 180 deg; joints [20.971, -63.816, 124.313, -156.232, 62.622, 78.552]
  MoveL 3343 to (-200, -20.47, 1.8) mm, rotated rx 0 ry 0 rz 180 deg; joints [20.971, -63.782, 124.319, -156.241, 62.659, 78.57]
  MoveL 3344 to (0, -20.47, 1.8) mm, rotated rx 0 ry 0 rz 180 deg; joints [18.129, -54.751, 108.376, -157.872, 55.693, 77.092]
  MoveL 3345 to (0, -19.87, 1.8) mm, rotated rx 0 ry 0 rz 180 deg; joints [18.129, -54.723, 108.382, -157.881, 55.725, 77.107]
  MoveL 3346 to (-200, -19.87, 1.8) mm, rotated rx 0 ry 0 rz 180 deg; joints [20.971, -63.748, 124.326, -156.249, 62.696, 78.589]
  MoveL 3347 to (-200, -19.27, 1.8) mm, rotated rx 0 ry 0 rz 180 deg; joints [20.971, -63.713, 124.332, -156.258, 62.734, 78.607]
  MoveL 3348 to (0, -19.27, 1.8) mm, rotated rx 0 ry 0 rz 180 deg; joints [18.129, -54.695, 108.388, -157.889, 55.756, 77.123]
  MoveL 3349 to (0, -18.67, 1.8) mm, rotated rx 0 ry 0 rz 180 deg; joints [18.129, -54.666, 108.394, -157.898, 55.788, 77.138]
  MoveL 3350 to (-200, -18.67, 1.8) mm, rotated rx 0 ry 0 rz 180 deg; joints [20.971, -63.679, 124.338, -156.266, 62.771, 78.625]
  MoveL 3351 to (-200, -18.07, 1.8) mm, rotated rx 0 ry 0 rz 180 deg; joints [20.971, -63.645, 124.344, -156.274, 62.808, 78.644]
  MoveL 3352 to (0, -18.07, 1.8) mm, rotated rx 0 ry 0 rz 180 deg; joints [18.129, -54.638, 108.4, -157.907, 55.82, 77.154]
  MoveL 3353 to (0, -17.47, 1.8) mm, rotated rx 0 ry 0 rz 180 deg; joints [18.129, -54.61, 108.405, -157.915, 55.851, 77.169]
  MoveL 3354 to (-200, -17.47, 1.8) mm, rotated rx 0 ry 0 rz 180 deg; joints [20.971, -63.611, 124.351, -156.283, 62.845, 78.662]
  MoveL 3355 to (-200, -16.87, 1.8) mm, rotated rx 0 ry 0 rz 180 deg; joints [20.971, -63.576, 124.357, -156.291, 62.882, 78.68]
  MoveL 3356 to (0, -16.87, 1.8) mm, rotated rx 0 ry 0 rz 180 deg; joints [18.129, -54.581, 108.411, -157.924, 55.883, 77.184]
  MoveL 3357 to (0, -16.27, 1.8) mm, rotated rx 0 ry 0 rz 180 deg; joints [18.129, -54.553, 108.417, -157.933, 55.914, 77.2]
  MoveL 3358 to (-200, -16.27, 1.8) mm, rotated rx 0 ry 0 rz 180 deg; joints [20.971, -63.542, 124.363, -156.299, 62.919, 78.699]
  MoveL 3359 to (-200, -15.67, 1.8) mm, rotated rx 0 ry 0 rz 180 deg; joints [20.971, -63.507, 124.369, -156.308, 62.957, 78.717]
  MoveL 3360 to (0, -15.67, 1.8) mm, rotated rx 0 ry 0 rz 180 deg; joints [18.129, -54.525, 108.423, -157.941, 55.946, 77.215]
  MoveL 3361 to (0, -15.07, 1.8) mm, rotated rx 0 ry 0 rz 180 deg; joints [18.129, -54.496, 108.428, -157.95, 55.977, 77.231]
  MoveL 3362 to (-200, -15.07, 1.8) mm, rotated rx 0 ry 0 rz 180 deg; joints [20.971, -63.473, 124.375, -156.316, 62.994, 78.735]
  MoveL 3363 to (-200, -14.47, 1.8) mm, rotated rx 0 ry 0 rz 180 deg; joints [20.971, -63.438, 124.381, -156.324, 63.031, 78.754]
  MoveL 3364 to (0, -14.47, 1.8) mm, rotated rx 0 ry 0 rz 180 deg; joints [18.129, -54.468, 108.434, -157.959, 56.009, 77.246]
  MoveL 3365 to (0, -13.87, 1.8) mm, rotated rx 0 ry 0 rz 180 deg; joints [18.129, -54.44, 108.439, -157.967, 56.04, 77.261]
  MoveL 3366 to (-200, -13.87, 1.8) mm, rotated rx 0 ry 0 rz 180 deg; joints [20.971, -63.404, 124.388, -156.333, 63.068, 78.772]
  MoveL 3367 to (-200, -13.27, 1.8) mm, rotated rx 0 ry 0 rz 180 deg; joints [20.971, -63.37, 124.394, -156.341, 63.105, 78.79]
  MoveL 3368 to (0, -13.27, 1.8) mm, rotated rx 0 ry 0 rz 180 deg; joints [18.129, -54.411, 108.445, -157.976, 56.072, 77.277]
  MoveL 3369 to (0, -12.67, 1.8) mm, rotated rx 0 ry 0 rz 180 deg; joints [18.129, -54.383, 108.45, -157.984, 56.103, 77.292]
  MoveL 3370 to (-200, -12.67, 1.8) mm, rotated rx 0 ry 0 rz 180 deg; joints [20.971, -63.335, 124.4, -156.349, 63.142, 78.808]
  MoveL 3371 to (-200, -12.07, 1.8) mm, rotated rx 0 ry 0 rz 180 deg; joints [20.971, -63.3, 124.406, -156.357, 63.179, 78.827]
  MoveL 3372 to (0, -12.07, 1.8) mm, rotated rx 0 ry 0 rz 180 deg; joints [18.129, -54.355, 108.456, -157.993, 56.134, 77.307]
  MoveL 3373 to (0, -11.47, 1.8) mm, rotated rx 0 ry 0 rz 180 deg; joints [18.129, -54.326, 108.461, -158.001, 56.166, 77.323]
  MoveL 3374 to (-200, -11.47, 1.8) mm, rotated rx 0 ry 0 rz 180 deg; joints [20.971, -63.266, 124.411, -156.366, 63.216, 78.845]
  MoveL 3375 to (-200, -10.87, 1.8) mm, rotated rx 0 ry 0 rz 180 deg; joints [20.971, -63.231, 124.417, -156.374, 63.253, 78.863]
  MoveL 3376 to (0, -10.87, 1.8) mm, rotated rx 0 ry 0 rz 180 deg; joints [18.129, -54.298, 108.467, -158.01, 56.197, 77.338]
  MoveL 3377 to (0, -10.27, 1.8) mm, rotated rx 0 ry 0 rz 180 deg; joints [18.129, -54.269, 108.472, -158.018, 56.229, 77.353]
  MoveL 3378 to (-200, -10.27, 1.8) mm, rotated rx 0 ry 0 rz 180 deg; joints [20.971, -63.197, 124.423, -156.382, 63.291, 78.881]
  MoveL 3379 to (-200, -9.67, 1.8) mm, rotated rx 0 ry 0 rz 180 deg; joints [20.971, -63.162, 124.429, -156.39, 63.328, 78.899]
  MoveL 3380 to (0, -9.67, 1.8) mm, rotated rx 0 ry 0 rz 180 deg; joints [18.129, -54.241, 108.478, -158.027, 56.26, 77.369]
  MoveL 3381 to (0, -9.07, 1.8) mm, rotated rx 0 ry 0 rz 180 deg; joints [18.129, -54.212, 108.483, -158.035, 56.292, 77.384]
  MoveL 3382 to (-200, -9.07, 1.8) mm, rotated rx 0 ry 0 rz 180 deg; joints [20.971, -63.127, 124.435, -156.398, 63.365, 78.917]
  MoveL 3383 to (-200, -8.47, 1.8) mm, rotated rx 0 ry 0 rz 180 deg; joints [20.971, -63.093, 124.441, -156.406, 63.402, 78.935]
  MoveL 3384 to (0, -8.47, 1.8) mm, rotated rx 0 ry 0 rz 180 deg; joints [18.129, -54.184, 108.488, -158.044, 56.323, 77.399]
  MoveL 3385 to (0, -7.87, 1.8) mm, rotated rx 0 ry 0 rz 180 deg; joints [18.129, -54.155, 108.494, -158.052, 56.354, 77.414]
  MoveL 3386 to (-200, -7.87, 1.8) mm, rotated rx 0 ry 0 rz 180 deg; joints [20.971, -63.058, 124.446, -156.414, 63.439, 78.953]
  MoveL 3387 to (-200, -7.27, 1.8) mm, rotated rx 0 ry 0 rz 180 deg; joints [20.971, -63.023, 124.452, -156.423, 63.476, 78.972]
  MoveL 3388 to (0, -7.27, 1.8) mm, rotated rx 0 ry 0 rz 180 deg; joints [18.129, -54.126, 108.499, -158.061, 56.386, 77.429]
  MoveL 3389 to (0, -6.67, 1.8) mm, rotated rx 0 ry 0 rz 180 deg; joints [18.129, -54.098, 108.504, -158.069, 56.417, 77.444]
  MoveL 3390 to (-200, -6.67, 1.8) mm, rotated rx 0 ry 0 rz 180 deg; joints [20.971, -62.989, 124.458, -156.431, 63.513, 78.99]
  MoveL 3391 to (-200, -6.07, 1.8) mm, rotated rx 0 ry 0 rz 180 deg; joints [20.971, -62.954, 124.463, -156.439, 63.55, 79.008]
  MoveL 3392 to (0, -6.07, 1.8) mm, rotated rx 0 ry 0 rz 180 deg; joints [18.129, -54.069, 108.509, -158.077, 56.448, 77.46]
  MoveL 3393 to (0, -5.47, 1.8) mm, rotated rx 0 ry 0 rz 180 deg; joints [18.129, -54.041, 108.514, -158.086, 56.48, 77.475]
  MoveL 3394 to (-200, -5.47, 1.8) mm, rotated rx 0 ry 0 rz 180 deg; joints [20.971, -62.919, 124.469, -156.447, 63.587, 79.026]
  MoveL 3395 to (-200, -4.87, 1.8) mm, rotated rx 0 ry 0 rz 180 deg; joints [20.971, -62.884, 124.475, -156.455, 63.624, 79.044]
  MoveL 3396 to (0, -4.87, 1.8) mm, rotated rx 0 ry 0 rz 180 deg; joints [18.129, -54.012, 108.519, -158.094, 56.511, 77.49]
  MoveL 3397 to (0, -4.27, 1.8) mm, rotated rx 0 ry 0 rz 180 deg; joints [18.129, -53.983, 108.525, -158.102, 56.542, 77.505]
  MoveL 3398 to (-200, -4.27, 1.8) mm, rotated rx 0 ry 0 rz 180 deg; joints [20.971, -62.85, 124.48, -156.463, 63.661, 79.062]
  MoveL 3399 to (-200, -3.67, 1.8) mm, rotated rx 0 ry 0 rz 180 deg; joints [20.971, -62.815, 124.486, -156.471, 63.698, 79.08]
  MoveL 3400 to (0, -3.67, 1.8) mm, rotated rx 0 ry 0 rz 180 deg; joints [18.129, -53.955, 108.53, -158.111, 56.574, 77.52]
  MoveL 3401 to (0, -3.07, 1.8) mm, rotated rx 0 ry 0 rz 180 deg; joints [18.129, -53.926, 108.535, -158.119, 56.605, 77.535]
  MoveL 3402 to (-200, -3.07, 1.8) mm, rotated rx 0 ry 0 rz 180 deg; joints [20.971, -62.78, 124.491, -156.479, 63.735, 79.098]
  MoveL 3403 to (-200, -2.47, 1.8) mm, rotated rx 0 ry 0 rz 180 deg; joints [20.971, -62.745, 124.497, -156.486, 63.772, 79.116]
  MoveL 3404 to (0, -2.47, 1.8) mm, rotated rx 0 ry 0 rz 180 deg; joints [18.129, -53.897, 108.54, -158.127, 56.636, 77.55]
  MoveL 3405 to (0, -1.87, 1.8) mm, rotated rx 0 ry 0 rz 180 deg; joints [18.129, -53.868, 108.545, -158.135, 56.668, 77.565]
  MoveL 3406 to (-200, -1.87, 1.8) mm, rotated rx 0 ry 0 rz 180 deg; joints [20.971, -62.71, 124.502, -156.494, 63.809, 79.133]
  MoveL 3407 to (-200, -1.27, 1.8) mm, rotated rx 0 ry 0 rz 180 deg; joints [20.971, -62.675, 124.507, -156.502, 63.846, 79.151]
  MoveL 3408 to (0, -1.27, 1.8) mm, rotated rx 0 ry 0 rz 180 deg; joints [18.129, -53.84, 108.55, -158.144, 56.699, 77.58]
  MoveL 3409 to (0, -0.67, 1.8) mm, rotated rx 0 ry 0 rz 180 deg; joints [18.129, -53.811, 108.555, -158.152, 56.73, 77.595]
  MoveL 3410 to (-200, -0.67, 1.8) mm, rotated rx 0 ry 0 rz 180 deg; joints [20.971, -62.64, 124.513, -156.51, 63.883, 79.169]
  MoveL 3411 to (-200, -0.07, 1.8) mm, rotated rx 0 ry 0 rz 180 deg; joints [20.971, -62.605, 124.518, -156.518, 63.92, 79.187]
  MoveL 3412 to (0, -0.07, 1.8) mm, rotated rx 0 ry 0 rz 180 deg; joints [18.129, -53.782, 108.56, -158.16, 56.761, 77.61]
  MoveL 3413 to (0, 0, 1.8) mm, rotated rx 0 ry 0 rz 180 deg; joints [18.129, -53.779, 108.56, -158.161, 56.765, 77.612]
  MoveL 3414 to (-200, 0, 1.8) mm, rotated rx 0 ry 0 rz 180 deg; joints [20.971, -62.601, 124.519, -156.519, 63.924, 79.189]
  MoveL 3415 to (-200, 0, 1.4) mm, rotated rx 0 ry 0 rz 180 deg; joints [20.988, -62.595, 124.507, -156.499, 63.923, 79.179]
  MoveL 3416 to (0, 0, 1.4) mm, rotated rx 0 ry 0 rz 180 deg; joints [18.144, -53.773, 108.549, -158.142, 56.764, 77.6]
  MoveL 3417 to (0, -0.6, 1.4) mm, rotated rx 0 ry 0 rz 180 deg; joints [18.144, -53.802, 108.544, -158.134, 56.732, 77.585]
  MoveL 3418 to (-200, -0.6, 1.4) mm, rotated rx 0 ry 0 rz 180 deg; joints [20.988, -62.63, 124.502, -156.491, 63.886, 79.161]
  MoveL 3419 to (-200, -1.2, 1.4) mm, rotated rx 0 ry 0 rz 180 deg; joints [20.988, -62.665, 124.496, -156.484, 63.849, 79.143]
  MoveL 3420 to (0, -1.2, 1.4) mm, rotated rx 0 ry 0 rz 180 deg; joints [18.144, -53.83, 108.539, -158.126, 56.701, 77.57]
  MoveL 3421 to (0, -1.8, 1.4) mm, rotated rx 0 ry 0 rz 180 deg; joints [18.144, -53.859, 108.534, -158.118, 56.67, 77.555]
  MoveL 3422 to (-200, -1.8, 1.4) mm, rotated rx 0 ry 0 rz 180 deg; joints [20.988, -62.7, 124.491, -156.476, 63.812, 79.125]
  MoveL 3423 to (-200, -2.4, 1.4) mm, rotated rx 0 ry 0 rz 180 deg; joints [20.988, -62.734, 124.486, -156.468, 63.775, 79.107]
  MoveL 3424 to (0, -2.4, 1.4) mm, rotated rx 0 ry 0 rz 180 deg; joints [18.144, -53.888, 108.529, -158.109, 56.638, 77.54]
  MoveL 3425 to (0, -3, 1.4) mm, rotated rx 0 ry 0 rz 180 deg; joints [18.144, -53.917, 108.524, -158.101, 56.607, 77.525]
  MoveL 3426 to (-200, -3, 1.4) mm, rotated rx 0 ry 0 rz 180 deg; joints [20.988, -62.769, 124.48, -156.46, 63.738, 79.089]
  MoveL 3427 to (-200, -3.6, 1.4) mm, rotated rx 0 ry 0 rz 180 deg; joints [20.988, -62.804, 124.475, -156.452, 63.701, 79.071]
  MoveL 3428 to (0, -3.6, 1.4) mm, rotated rx 0 ry 0 rz 180 deg; joints [18.144, -53.945, 108.519, -158.093, 56.576, 77.51]
  MoveL 3429 to (0, -4.2, 1.4) mm, rotated rx 0 ry 0 rz 180 deg; joints [18.144, -53.974, 108.514, -158.084, 56.545, 77.495]
  MoveL 3430 to (-200, -4.2, 1.4) mm, rotated rx 0 ry 0 rz 180 deg; joints [20.988, -62.839, 124.469, -156.444, 63.664, 79.053]
  MoveL 3431 to (-200, -4.8, 1.4) mm, rotated rx 0 ry 0 rz 180 deg; joints [20.988, -62.874, 124.464, -156.436, 63.627, 79.035]
  MoveL 3432 to (0, -4.8, 1.4) mm, rotated rx 0 ry 0 rz 180 deg; joints [18.144, -54.003, 108.509, -158.076, 56.513, 77.48]
  MoveL 3433 to (0, -5.4, 1.4) mm, rotated rx 0 ry 0 rz 180 deg; joints [18.144, -54.031, 108.504, -158.068, 56.482, 77.464]
  MoveL 3434 to (-200, -5.4, 1.4) mm, rotated rx 0 ry 0 rz 180 deg; joints [20.988, -62.909, 124.458, -156.428, 63.59, 79.017]
  MoveL 3435 to (-200, -6, 1.4) mm, rotated rx 0 ry 0 rz 180 deg; joints [20.988, -62.943, 124.453, -156.42, 63.553, 78.999]
  MoveL 3436 to (0, -6, 1.4) mm, rotated rx 0 ry 0 rz 180 deg; joints [18.144, -54.06, 108.499, -158.059, 56.451, 77.449]
  MoveL 3437 to (0, -6.6, 1.4) mm, rotated rx 0 ry 0 rz 180 deg; joints [18.144, -54.088, 108.493, -158.051, 56.419, 77.434]
  MoveL 3438 to (-200, -6.6, 1.4) mm, rotated rx 0 ry 0 rz 180 deg; joints [20.988, -62.978, 124.447, -156.412, 63.516, 78.981]
  MoveL 3439 to (-200, -7.2, 1.4) mm, rotated rx 0 ry 0 rz 180 deg; joints [20.988, -63.013, 124.441, -156.404, 63.479, 78.963]
  MoveL 3440 to (0, -7.2, 1.4) mm, rotated rx 0 ry 0 rz 180 deg; joints [18.144, -54.117, 108.488, -158.043, 56.388, 77.419]
  MoveL 3441 to (0, -7.8, 1.4) mm, rotated rx 0 ry 0 rz 180 deg; joints [18.144, -54.146, 108.483, -158.034, 56.356, 77.404]
  MoveL 3442 to (-200, -7.8, 1.4) mm, rotated rx 0 ry 0 rz 180 deg; joints [20.988, -63.048, 124.435, -156.396, 63.442, 78.945]
  MoveL 3443 to (-200, -8.4, 1.4) mm, rotated rx 0 ry 0 rz 180 deg; joints [20.988, -63.082, 124.43, -156.388, 63.405, 78.927]
  MoveL 3444 to (0, -8.4, 1.4) mm, rotated rx 0 ry 0 rz 180 deg; joints [18.144, -54.174, 108.478, -158.026, 56.325, 77.389]
  MoveL 3445 to (0, -9, 1.4) mm, rotated rx 0 ry 0 rz 180 deg; joints [18.144, -54.203, 108.472, -158.017, 56.294, 77.373]
  MoveL 3446 to (-200, -9, 1.4) mm, rotated rx 0 ry 0 rz 180 deg; joints [20.988, -63.117, 124.424, -156.379, 63.368, 78.909]
  MoveL 3447 to (-200, -9.6, 1.4) mm, rotated rx 0 ry 0 rz 180 deg; joints [20.988, -63.152, 124.418, -156.371, 63.331, 78.891]
  MoveL 3448 to (0, -9.6, 1.4) mm, rotated rx 0 ry 0 rz 180 deg; joints [18.144, -54.231, 108.467, -158.009, 56.262, 77.358]
  MoveL 3449 to (0, -10.2, 1.4) mm, rotated rx 0 ry 0 rz 180 deg; joints [18.144, -54.26, 108.462, -158, 56.231, 77.343]
  MoveL 3450 to (-200, -10.2, 1.4) mm, rotated rx 0 ry 0 rz 180 deg; joints [20.988, -63.186, 124.412, -156.363, 63.294, 78.873]
  MoveL 3451 to (-200, -10.8, 1.4) mm, rotated rx 0 ry 0 rz 180 deg; joints [20.988, -63.221, 124.406, -156.355, 63.257, 78.854]
  MoveL 3452 to (0, -10.8, 1.4) mm, rotated rx 0 ry 0 rz 180 deg; joints [18.144, -54.288, 108.456, -157.992, 56.2, 77.328]
  MoveL 3453 to (0, -11.4, 1.4) mm, rotated rx 0 ry 0 rz 180 deg; joints [18.144, -54.317, 108.451, -157.983, 56.168, 77.312]
  MoveL 3454 to (-200, -11.4, 1.4) mm, rotated rx 0 ry 0 rz 180 deg; joints [20.988, -63.255, 124.401, -156.347, 63.219, 78.836]
  MoveL 3455 to (-200, -12, 1.4) mm, rotated rx 0 ry 0 rz 180 deg; joints [20.988, -63.29, 124.395, -156.339, 63.182, 78.818]
  MoveL 3456 to (0, -12, 1.4) mm, rotated rx 0 ry 0 rz 180 deg; joints [18.144, -54.345, 108.445, -157.975, 56.137, 77.297]
  MoveL 3457 to (0, -12.6, 1.4) mm, rotated rx 0 ry 0 rz 180 deg; joints [18.144, -54.374, 108.44, -157.966, 56.105, 77.282]
  MoveL 3458 to (-200, -12.6, 1.4) mm, rotated rx 0 ry 0 rz 180 deg; joints [20.988, -63.324, 124.389, -156.33, 63.145, 78.8]
  MoveL 3459 to (-200, -13.2, 1.4) mm, rotated rx 0 ry 0 rz 180 deg; joints [20.988, -63.359, 124.383, -156.322, 63.108, 78.782]
  MoveL 3460 to (0, -13.2, 1.4) mm, rotated rx 0 ry 0 rz 180 deg; joints [18.144, -54.402, 108.434, -157.958, 56.074, 77.266]
  MoveL 3461 to (0, -13.8, 1.4) mm, rotated rx 0 ry 0 rz 180 deg; joints [18.144, -54.43, 108.429, -157.949, 56.042, 77.251]
  MoveL 3462 to (-200, -13.8, 1.4) mm, rotated rx 0 ry 0 rz 180 deg; joints [20.988, -63.393, 124.377, -156.314, 63.071, 78.763]
  MoveL 3463 to (-200, -14.4, 1.4) mm, rotated rx 0 ry 0 rz 180 deg; joints [20.988, -63.428, 124.371, -156.306, 63.034, 78.745]
  MoveL 3464 to (0, -14.4, 1.4) mm, rotated rx 0 ry 0 rz 180 deg; joints [18.144, -54.459, 108.423, -157.941, 56.011, 77.236]
  MoveL 3465 to (0, -15, 1.4) mm, rotated rx 0 ry 0 rz 180 deg; joints [18.144, -54.487, 108.418, -157.932, 55.979, 77.22]
  MoveL 3466 to (-200, -15, 1.4) mm, rotated rx 0 ry 0 rz 180 deg; joints [20.988, -63.462, 124.365, -156.297, 62.997, 78.727]
  MoveL 3467 to (-200, -15.6, 1.4) mm, rotated rx 0 ry 0 rz 180 deg; joints [20.988, -63.497, 124.358, -156.289, 62.96, 78.708]
  MoveL 3468 to (0, -15.6, 1.4) mm, rotated rx 0 ry 0 rz 180 deg; joints [18.144, -54.515, 108.412, -157.923, 55.948, 77.205]
  MoveL 3469 to (0, -16.2, 1.4) mm, rotated rx 0 ry 0 rz 180 deg; joints [18.144, -54.544, 108.406, -157.915, 55.916, 77.189]
  MoveL 3470 to (-200, -16.2, 1.4) mm, rotated rx 0 ry 0 rz 180 deg; joints [20.988, -63.531, 124.352, -156.281, 62.923, 78.69]
  MoveL 3471 to (-200, -16.8, 1.4) mm, rotated rx 0 ry 0 rz 180 deg; joints [20.988, -63.565, 124.346, -156.272, 62.886, 78.672]
  MoveL 3472 to (0, -16.8, 1.4) mm, rotated rx 0 ry 0 rz 180 deg; joints [18.144, -54.572, 108.401, -157.906, 55.885, 77.174]
  MoveL 3473 to (0, -17.4, 1.4) mm, rotated rx 0 ry 0 rz 180 deg; joints [18.144, -54.6, 108.395, -157.897, 55.853, 77.159]
  MoveL 3474 to (-200, -17.4, 1.4) mm, rotated rx 0 ry 0 rz 180 deg; joints [20.988, -63.6, 124.34, -156.264, 62.848, 78.653]
  MoveL 3475 to (-200, -18, 1.4) mm, rotated rx 0 ry 0 rz 180 deg; joints [20.988, -63.634, 124.334, -156.256, 62.811, 78.635]
  MoveL 3476 to (0, -18, 1.4) mm, rotated rx 0 ry 0 rz 180 deg; joints [18.144, -54.629, 108.389, -157.889, 55.822, 77.143]
  MoveL 3477 to (0, -18.6, 1.4) mm, rotated rx 0 ry 0 rz 180 deg; joints [18.144, -54.657, 108.383, -157.88, 55.79, 77.128]
  MoveL 3478 to (-200, -18.6, 1.4) mm, rotated rx 0 ry 0 rz 180 deg; joints [20.988, -63.669, 124.327, -156.247, 62.774, 78.617]
  MoveL 3479 to (-200, -19.2, 1.4) mm, rotated rx 0 ry 0 rz 180 deg; joints [20.988, -63.703, 124.321, -156.239, 62.737, 78.598]
  MoveL 3480 to (0, -19.2, 1.4) mm, rotated rx 0 ry 0 rz 180 deg; joints [18.144, -54.685, 108.378, -157.871, 55.759, 77.112]
  MoveL 3481 to (0, -19.8, 1.4) mm, rotated rx 0 ry 0 rz 180 deg; joints [18.144, -54.713, 108.372, -157.862, 55.727, 77.097]
  MoveL 3482 to (-200, -19.8, 1.4) mm, rotated rx 0 ry 0 rz 180 deg; joints [20.988, -63.737, 124.315, -156.23, 62.7, 78.58]
  MoveL 3483 to (-200, -20.4, 1.4) mm, rotated rx 0 ry 0 rz 180 deg; joints [20.988, -63.771, 124.308, -156.222, 62.663, 78.561]
  MoveL 3484 to (0, -20.4, 1.4) mm, rotated rx 0 ry 0 rz 180 deg; joints [18.144, -54.742, 108.366, -157.854, 55.696, 77.081]
  MoveL 3485 to (0, -21, 1.4) mm, rotated rx 0 ry 0 rz 180 deg; joints [18.144, -54.77, 108.36, -157.845, 55.664, 77.065]
  MoveL 3486 to (-200, -21, 1.4) mm, rotated rx 0 ry 0 rz 180 deg; joints [20.988, -63.806, 124.302, -156.213, 62.625, 78.543]
  MoveL 3487 to (-200, -21.6, 1.4) mm, rotated rx 0 ry 0 rz 180 deg; joints [20.988, -63.84, 124.296, -156.205, 62.588, 78.525]
  MoveL 3488 to (0, -21.6, 1.4) mm, rotated rx 0 ry 0 rz 180 deg; joints [18.144, -54.798, 108.354, -157.836, 55.633, 77.05]
  MoveL 3489 to (0, -22.2, 1.4) mm, rotated rx 0 ry 0 rz 180 deg; joints [18.144, -54.826, 108.348, -157.827, 55.601, 77.034]
  MoveL 3490 to (-200, -22.2, 1.4) mm, rotated rx 0 ry 0 rz 180 deg; joints [20.988, -63.874, 124.289, -156.196, 62.551, 78.506]
  MoveL 3491 to (-200, -22.8, 1.4) mm, rotated rx 0 ry 0 rz 180 deg; joints [20.988, -63.908, 124.283, -156.188, 62.514, 78.488]
  MoveL 3492 to (0, -22.8, 1.4) mm, rotated rx 0 ry 0 rz 180 deg; joints [18.144, -54.854, 108.342, -157.819, 55.569, 77.019]
  MoveL 3493 to (0, -23.4, 1.4) mm, rotated rx 0 ry 0 rz 180 deg; joints [18.144, -54.882, 108.336, -157.81, 55.538, 77.003]
  MoveL 3494 to (-200, -23.4, 1.4) mm, rotated rx 0 ry 0 rz 180 deg; joints [20.988, -63.942, 124.276, -156.179, 62.477, 78.469]
  MoveL 3495 to (-200, -24, 1.4) mm, rotated rx 0 ry 0 rz 180 deg; joints [20.988, -63.976, 124.269, -156.171, 62.439, 78.451]
  MoveL 3496 to (0, -24, 1.4) mm, rotated rx 0 ry 0 rz 180 deg; joints [18.144, -54.91, 108.33, -157.801, 55.506, 76.987]
  MoveL 3497 to (0, -24.6, 1.4) mm, rotated rx 0 ry 0 rz 180 deg; joints [18.144, -54.938, 108.324, -157.792, 55.475, 76.972]
  MoveL 3498 to (-200, -24.6, 1.4) mm, rotated rx 0 ry 0 rz 180 deg; joints [20.988, -64.01, 124.263, -156.162, 62.402, 78.432]
  MoveL 3499 to (-200, -25.2, 1.4) mm, rotated rx 0 ry 0 rz 180 deg; joints [20.988, -64.045, 124.256, -156.154, 62.365, 78.413]
  MoveL 3500 to (0, -25.2, 1.4) mm, rotated rx 0 ry 0 rz 180 deg; joints [18.144, -54.966, 108.318, -157.783, 55.443, 76.956]
  MoveL 3501 to (0, -25.8, 1.4) mm, rotated rx 0 ry 0 rz 180 deg; joints [18.144, -54.994, 108.312, -157.774, 55.411, 76.94]
  MoveL 3502 to (-200, -25.8, 1.4) mm, rotated rx 0 ry 0 rz 180 deg; joints [20.988, -64.079, 124.25, -156.145, 62.328, 78.395]
  MoveL 3503 to (-200, -26.4, 1.4) mm, rotated rx 0 ry 0 rz 180 deg; joints [20.988, -64.113, 124.243, -156.136, 62.29, 78.376]
  MoveL 3504 to (0, -26.4, 1.4) mm, rotated rx 0 ry 0 rz 180 deg; joints [18.144, -55.022, 108.306, -157.765, 55.38, 76.925]
  MoveL 3505 to (0, -27, 1.4) mm, rotated rx 0 ry 0 rz 180 deg; joints [18.144, -55.05, 108.299, -157.756, 55.348, 76.909]
  MoveL 3506 to (-200, -27, 1.4) mm, rotated rx 0 ry 0 rz 180 deg; joints [20.988, -64.147, 124.236, -156.128, 62.253, 78.358]
  MoveL 3507 to (-200, -27.6, 1.4) mm, rotated rx 0 ry 0 rz 180 deg; joints [20.988, -64.181, 124.229, -156.119, 62.216, 78.339]
  MoveL 3508 to (0, -27.6, 1.4) mm, rotated rx 0 ry 0 rz 180 deg; joints [18.144, -55.078, 108.293, -157.747, 55.316, 76.893]
  MoveL 3509 to (0, -28.2, 1.4) mm, rotated rx 0 ry 0 rz 180 deg; joints [18.144, -55.106, 108.287, -157.738, 55.285, 76.877]
  MoveL 3510 to (-200, -28.2, 1.4) mm, rotated rx 0 ry 0 rz 180 deg; joints [20.988, -64.215, 124.223, -156.11, 62.179, 78.32]
  MoveL 3511 to (-200, -28.8, 1.4) mm, rotated rx 0 ry 0 rz 180 deg; joints [20.988, -64.249, 124.216, -156.101, 62.141, 78.302]
  MoveL 3512 to (0, -28.8, 1.4) mm, rotated rx 0 ry 0 rz 180 deg; joints [18.144, -55.134, 108.281, -157.729, 55.253, 76.862]
  MoveL 3513 to (0, -29.4, 1.4) mm, rotated rx 0 ry 0 rz 180 deg; joints [18.144, -55.162, 108.274, -157.72, 55.221, 76.846]
  MoveL 3514 to (-200, -29.4, 1.4) mm, rotated rx 0 ry 0 rz 180 deg; joints [20.988, -64.282, 124.209, -156.093, 62.104, 78.283]
  MoveL 3515 to (-200, -30, 1.4) mm, rotated rx 0 ry 0 rz 180 deg; joints [20.988, -64.316, 124.202, -156.084, 62.067, 78.264]
  MoveL 3516 to (0, -30, 1.4) mm, rotated rx 0 ry 0 rz 180 deg; joints [18.144, -55.19, 108.268, -157.711, 55.19, 76.83]
  MoveL 3517 to (0, -30.6, 1.41) mm, rotated rx 2.53 ry 0 rz 180 deg; joints [18.058, -55.978, 108.147, -157.569, 54.329, 78.993]
  MoveL 3518 to (-200, -30.6, 1.41) mm, rotated rx 2.53 ry 0 rz 180 deg; joints [20.891, -65.27, 124.068, -155.952, 61.053, 80.341]
  MoveL 3519 to (-200, -31.2, 1.45) mm, rotated rx 5.06 ry 0 rz 180 deg; joints [20.763, -66.214, 123.932, -155.846, 60.039, 82.432]
  MoveL 3520 to (0, -31.2, 1.45) mm, rotated rx 5.06 ry 0 rz 180 deg; joints [17.945, -56.76, 108.026, -157.453, 53.468, 81.174]
  MoveL 3521 to (0, -31.8, 1.52) mm, rotated rx 7.58 ry 0 rz 180 deg; joints [17.806, -57.532, 107.904, -157.364, 52.608, 83.373]
  MoveL 3522 to (-200, -31.8, 1.52) mm, rotated rx 7.58 ry 0 rz 180 deg; joints [20.605, -67.148, 123.794, -155.767, 59.027, 84.541]
  MoveL 3523 to (-200, -32.39, 1.61) mm, rotated rx 10.11 ry 0 rz 180 deg; joints [20.416, -68.069, 123.656, -155.716, 58.018, 86.671]
  MoveL 3524 to (0, -32.39, 1.61) mm, rotated rx 10.11 ry 0 rz 180 deg; joints [17.639, -58.296, 107.781, -157.303, 51.75, 85.594]
  MoveL 3525 to (0, -32.98, 1.73) mm, rotated rx 12.64 ry 0 rz 180 deg; joints [17.445, -59.049, 107.66, -157.273, 50.894, 87.84]
  MoveL 3526 to (-200, -32.98, 1.73) mm, rotated rx 12.64 ry 0 rz 180 deg; joints [20.197, -68.977, 123.517, -155.694, 57.012, 88.824]
  MoveL 3527 to (-200, -33.56, 1.87) mm, rotated rx 15.17 ry 0 rz 180 deg; joints [19.948, -69.87, 123.378, -155.703, 56.011, 91.003]
  MoveL 3528 to (0, -33.56, 1.87) mm, rotated rx 15.17 ry 0 rz 180 deg; joints [17.225, -59.789, 107.539, -157.274, 50.042, 90.112]
  MoveL 3529 to (0, -34.13, 2.04) mm, rotated rx 17.69 ry 0 rz 180 deg; joints [16.978, -60.517, 107.419, -157.308, 49.196, 92.411]
  MoveL 3530 to (-200, -34.13, 2.04) mm, rotated rx 17.69 ry 0 rz 180 deg; joints [19.668, -70.746, 123.24, -155.746, 55.018, 93.21]
  MoveL 3531 to (-200, -34.7, 2.24) mm, rotated rx 20.22 ry 0 rz 180 deg; joints [19.359, -71.605, 123.103, -155.822, 54.031, 95.45]
  MoveL 3532 to (0, -34.7, 2.24) mm, rotated rx 20.22 ry 0 rz 180 deg; joints [16.706, -61.23, 107.301, -157.377, 48.357, 94.744]
  MoveL 3533 to (0, -35.26, 2.46) mm, rotated rx 22.75 ry 0 rz 180 deg; joints [16.408, -61.928, 107.185, -157.482, 47.525, 97.11]
  MoveL 3534 to (-200, -35.26, 2.46) mm, rotated rx 22.75 ry 0 rz 180 deg; joints [19.02, -72.445, 122.968, -155.935, 53.054, 97.724]
  MoveL 3535 to (-200, -35.81, 2.7) mm, rotated rx 25.28 ry 0 rz 180 deg; joints [18.652, -73.264, 122.835, -156.086, 52.088, 100.037]
  MoveL 3536 to (0, -35.81, 2.7) mm, rotated rx 25.28 ry 0 rz 180 deg; joints [16.084, -62.61, 107.072, -157.625, 46.703, 99.514]
  MoveL 3537 to (0, -36.34, 2.97) mm, rotated rx 27.8 ry 0 rz 180 deg; joints [15.736, -63.274, 106.962, -157.809, 45.892, 101.955]
  MoveL 3538 to (-200, -36.34, 2.97) mm, rotated rx 27.8 ry 0 rz 180 deg; joints [18.255, -74.062, 122.704, -156.278, 51.134, 102.389]
  MoveL 3539 to (-200, -36.87, 3.26) mm, rotated rx 30.33 ry 0 rz 180 deg; joints [17.829, -74.837, 122.578, -156.512, 50.194, 104.786]
  MoveL 3540 to (0, -36.87, 3.26) mm, rotated rx 30.33 ry 0 rz 180 deg; joints [15.363, -63.919, 106.855, -158.034, 45.094, 104.44]
  MoveL 3541 to (0, -37.38, 3.58) mm, rotated rx 32.86 ry 0 rz 180 deg; joints [14.966, -64.545, 106.753, -158.304, 44.309, 106.969]
  MoveL 3542 to (-200, -37.38, 3.58) mm, rotated rx 32.86 ry 0 rz 180 deg; joints [17.376, -75.588, 122.455, -156.79, 49.27, 107.23]
  MoveL 3543 to (-200, -37.88, 3.91) mm, rotated rx 35.39 ry 0 rz 180 deg; joints [16.895, -76.315, 122.338, -157.116, 48.363, 109.724]
  MoveL 3544 to (0, -37.88, 3.91) mm, rotated rx 35.39 ry 0 rz 180 deg; joints [14.545, -65.15, 106.656, -158.619, 43.541, 109.545]
  MoveL 3545 to (0, -38.36, 4.27) mm, rotated rx 37.92 ry 0 rz 180 deg; joints [14.102, -65.733, 106.564, -158.982, 42.791, 112.17]
  MoveL 3546 to (-200, -38.36, 4.27) mm, rotated rx 37.92 ry 0 rz 180 deg; joints [16.388, -77.015, 122.225, -157.491, 47.477, 112.27]
  MoveL 3547 to (-200, -38.82, 4.65) mm, rotated rx 40.44 ry 0 rz 180 deg; joints [15.855, -77.689, 122.119, -157.918, 46.612, 114.872]
  MoveL 3548 to (0, -38.82, 4.65) mm, rotated rx 40.44 ry 0 rz 180 deg; joints [13.636, -66.294, 106.478, -159.395, 42.06, 114.847]
  MoveL 3549 to (0, -39.27, 5.05) mm, rotated rx 42.97 ry 0 rz 180 deg; joints [13.15, -66.832, 106.398, -159.859, 41.351, 117.578]
  MoveL 3550 to (-200, -39.27, 5.05) mm, rotated rx 42.97 ry 0 rz 180 deg; joints [15.296, -78.334, 122.02, -158.399, 45.771, 117.533]
  MoveL 3551 to (-200, -39.7, 5.47) mm, rotated rx 45.5 ry 0 rz 180 deg; joints [14.712, -78.951, 121.928, -158.935, 44.957, 120.254]
  MoveL 3552 to (0, -39.7, 5.47) mm, rotated rx 45.5 ry 0 rz 180 deg; joints [12.642, -67.346, 106.325, -160.376, 40.666, 120.366]
  MoveL 3553 to (0, -40.11, 5.91) mm, rotated rx 48.03 ry 0 rz 180 deg; joints [12.115, -67.835, 106.26, -160.946, 40.006, 123.209]
  MoveL 3554 to (-200, -40.11, 5.91) mm, rotated rx 48.03 ry 0 rz 180 deg; joints [14.105, -79.537, 121.844, -159.529, 44.172, 123.037]
  MoveL 3555 to (-200, -40.5, 6.36) mm, rotated rx 50.55 ry 0 rz 180 deg; joints [13.475, -80.092, 121.768, -160.182, 43.419, 125.886]
  MoveL 3556 to (0, -40.5, 6.36) mm, rotated rx 50.55 ry 0 rz 180 deg; joints [11.568, -68.298, 106.202, -161.573, 39.375, 126.112]
  MoveL 3557 to (0, -40.87, 6.83) mm, rotated rx 53.08 ry 0 rz 180 deg; joints [11.004, -68.734, 106.153, -162.255, 38.775, 129.075]
  MoveL 3558 to (-200, -40.87, 6.83) mm, rotated rx 53.08 ry 0 rz 180 deg; joints [12.824, -80.616, 121.702, -160.895, 42.699, 128.801]
  MoveL 3559 to (-200, -41.22, 7.32) mm, rotated rx 55.61 ry 0 rz 180 deg; joints [12.152, -81.107, 121.645, -161.67, 42.017, 131.783]
  MoveL 3560 to (0, -41.22, 7.32) mm, rotated rx 55.61 ry 0 rz 180 deg; joints [10.422, -69.143, 106.112, -162.993, 38.207, 132.097]
  MoveL 3561 to (0, -41.55, 7.82) mm, rotated rx 58.14 ry 0 rz 180 deg; joints [9.825, -69.524, 106.081, -163.787, 37.675, 135.178]
  MoveL 3562 to (-200, -41.55, 7.82) mm, rotated rx 58.14 ry 0 rz 180 deg; joints [11.461, -81.565, 121.599, -162.506, 41.375, 134.831]
  MoveL 3563 to (-200, -41.86, 8.34) mm, rotated rx 60.67 ry 0 rz 180 deg; joints [10.751, -81.988, 121.563, -163.403, 40.776, 137.947]
  MoveL 3564 to (0, -41.86, 8.34) mm, rotated rx 60.67 ry 0 rz 180 deg; joints [9.213, -69.877, 106.059, -164.637, 37.181, 138.318]
  MoveL 3565 to (0, -42.14, 8.87) mm, rotated rx 63.19 ry 0 rz 180 deg; joints [8.588, -70.201, 106.047, -165.54, 36.726, 141.516]
  MoveL 3566 to (-200, -42.14, 8.87) mm, rotated rx 63.19 ry 0 rz 180 deg; joints [10.025, -82.377, 121.538, -164.361, 40.223, 141.129]
  MoveL 3567 to (-200, -42.4, 9.41) mm, rotated rx 65.72 ry 0 rz 180 deg; joints [9.284, -82.73, 121.524, -165.376, 39.719, 144.374]
  MoveL 3568 to (0, -42.4, 9.41) mm, rotated rx 65.72 ry 0 rz 180 deg; joints [7.95, -70.495, 106.045, -166.495, 36.314, 144.769]
  MoveL 3569 to (0, -42.63, 9.96) mm, rotated rx 68.25 ry 0 rz 180 deg; joints [7.301, -70.758, 106.053, -167.498, 35.946, 148.072]
  MoveL 3570 to (-200, -42.63, 9.96) mm, rotated rx 68.25 ry 0 rz 180 deg; joints [8.53, -83.047, 121.523, -166.447, 39.266, 147.678]
  MoveL 3571 to (-200, -42.84, 10.52) mm, rotated rx 70.78 ry 0 rz 180 deg; joints [7.763, -83.328, 121.533, -167.57, 38.868, 151.04]
  MoveL 3572 to (0, -42.84, 10.52) mm, rotated rx 70.78 ry 0 rz 180 deg; joints [6.642, -70.991, 106.072, -168.547, 35.625, 151.425]
  MoveL 3573 to (0, -43.03, 11.09) mm, rotated rx 73.31 ry 0 rz 180 deg; joints [5.975, -71.193, 106.102, -169.636, 35.353, 154.821]
  MoveL 3574 to (-200, -43.03, 11.09) mm, rotated rx 73.31 ry 0 rz 180 deg; joints [6.985, -83.571, 121.556, -168.741, 38.527, 154.453]
  MoveL 3575 to (-200, -43.19, 11.67) mm, rotated rx 75.83 ry 0 rz 180 deg; joints [6.199, -83.776, 121.591, -169.954, 38.245, 157.912]
  MoveL 3576 to (0, -43.19, 11.67) mm, rotated rx 75.83 ry 0 rz 180 deg; joints [5.301, -71.363, 106.143, -170.761, 35.131, 158.256]
  MoveL 3577 to (0, -43.32, 12.26) mm, rotated rx 78.36 ry 0 rz 180 deg; joints [4.622, -71.502, 106.194, -171.916, 34.961, 161.721]
  MoveL 3578 to (-200, -43.32, 12.26) mm, rotated rx 78.36 ry 0 rz 180 deg; joints [5.406, -83.943, 121.639, -171.202, 38.025, 161.409]
  MoveL 3579 to (-200, -43.43, 12.85) mm, rotated rx 80.89 ry 0 rz 180 deg; joints [4.608, -84.071, 121.699, -172.48, 37.867, 164.939]
  MoveL 3580 to (0, -43.43, 12.85) mm, rotated rx 80.89 ry 0 rz 180 deg; joints [3.938, -71.608, 106.257, -173.096, 34.844, 165.213]
  MoveL 3581 to (0, -43.51, 13.44) mm, rotated rx 83.42 ry 0 rz 180 deg; joints [3.253, -71.681, 106.33, -174.292, 34.782, 168.723]
  MoveL 3582 to (-200, -43.51, 13.44) mm, rotated rx 83.42 ry 0 rz 180 deg; joints [3.806, -84.161, 121.772, -173.779, 37.775, 168.492]
  MoveL 3583 to (-200, -43.57, 14.04) mm, rotated rx 85.94 ry 0 rz 180 deg; joints [3.003, -84.211, 121.858, -175.091, 37.749, 172.059]
  MoveL 3584 to (0, -43.57, 14.04) mm, rotated rx 85.94 ry 0 rz 180 deg; joints [2.566, -71.722, 106.414, -175.498, 34.775, 172.244]
  MoveL 3585 to (0, -43.59, 14.64) mm, rotated rx 88.47 ry 0 rz 180 deg; joints [1.88, -71.73, 106.508, -176.706, 34.823, 175.766]
  MoveL 3586 to (-200, -43.59, 14.64) mm, rotated rx 88.47 ry 0 rz 180 deg; joints [2.201, -84.222, 121.956, -176.407, 37.788, 175.63]
  MoveL 3587 to (-200, -43.6, 15.24) mm, rotated rx 90 ry 0 rz 180 deg; joints [1.705, -84.209, 122.021, -177.221, 37.844, 177.805]
  MoveL 3588 to (0, -43.6, 15.24) mm, rotated rx 90 ry 0 rz 180 deg; joints [1.456, -71.719, 106.571, -177.453, 34.878, 177.91]
  MoveL 3589 to (0, -43.6, 15.84) mm, rotated rx 90 ry 0 rz 180 deg; joints [1.431, -71.72, 106.572, -177.497, 34.878, 177.946]
  MoveL 3590 to (-200, -43.6, 15.84) mm, rotated rx 90 ry 0 rz 180 deg; joints [1.675, -84.21, 122.022, -177.269, 37.844, 177.843]
  MoveL 3591 to (-200, -43.6, 16.44) mm, rotated rx 90 ry 0 rz 180 deg; joints [1.646, -84.212, 122.024, -177.317, 37.843, 177.88]
